(* IEC 61131-3 sources: daoli-st-library/DL_MathData (part 31) *)

(* ---- FC_DL_CalcDistance3D.st ---- *)
(*==============================================================================
 * 组件名称 (Component)  : FC_DL_CalcDistance3D
 * 所属子库 (Sublibrary) : DL_MathData
 * 当前版本 (Version)    : 1.0.0
 * 分类     (Category)   : 几何计算函数（Function · Math / Pure function）
 * 兼容性   (Platform)   : CODESYS 3.5 / TwinCAT 3 / 汇川 InoProShop / Machine Expert
 *                         仅依赖 Standard.library（SQRT / ABS / MAX），零厂商方言
 * 功能描述 (Function)   : 计算两点之间的三维欧氏距离，附带非有限值防护、
 *                         大数溢出缩放保护与三个分量差诊断输出。
 *                         平面（二维）距离不另设组件：把两个端点的 Z 坐标
 *                         同时填 0.0 即为其退化情形，规格明确禁止为凑数拆变体。
 *                         全程无内部状态，可任意频次调用。
 *
 * 【引脚契约 / Pin contract】
 *   输入 fX1 / fY1 / fZ1 : REAL — 点 1 的 X / Y / Z 坐标 [mm]，量程 ±1.0E6，
 *                                  平面场景把两个 Z 都填 0.0；
 *   输入 fX2 / fY2 / fZ2 : REAL — 点 2 的 X / Y / Z 坐标 [mm]，量程同上；
 *   输出 bValid          : BOOL — 六个输入全部有限（非 NaN、非无穷）= TRUE；
 *   输出 bSaturated      : BOOL — 本次计算进入大数缩放分支（结果仍然有效，
 *                                  但已落在置信区间，提示调用方复核量纲）；
 *   输出 fDeltaX/Y/Z     : REAL — 三个分量差 [mm]，便于现场诊断「差在哪个轴」；
 *   输出 uErrorId        : UDINT — 事件码，0 = 无。本件全部码为信息级。
 *   返回  值             : REAL — 距离 [mm]，恒非负；输入非法时返回 0.0。
 *
 * 【算法分步 / Algorithm steps（写死，防实现漂移）】
 *   ① 有限性闸门：六个输入任一非有限 → bValid FALSE、返回 0.0、置 0122 后早退。
 *      刻意**不返回 NaN**：NaN 会沿调用链污染下游滤波、比较与统计（历史教训）；
 *   ② 分量差：dX = X2 − X1（同 Y、Z），同时作为诊断输出；
 *   ③ 比例因子：fScale = MAX(|dX|, |dY|, |dZ|)，取最大分量作为量级基准；
 *   ④ 分支一（常规）：fScale 小于缩放阈值 → 直接 SQRT(dX² + dY² + dZ²)；
 *   ⑤ 分支二（缩放）：fScale 超阈值 → SQRT((dX/fScale)² + (dY/fScale)² +
 *      (dZ/fScale)²) × fScale。归一后每一项绝对值不超过 1，平方和不超过 3，
 *      彻底规避「大数先平方再开方」的中间溢出，结果为同一数学量的稳定写法；
 *   ⑥ 退化：三个分量差全为零（同一点）→ 返回 0.0 且不置任何码，因为距离为 0
 *      是合法结果而不是异常；
 *   ⑦ 后置守卫：最终结果非有限时（理论上不可达，防御性兜底）返回 0.0 并置 0122。
 *
 * 【数值安全 / Numeric safety】
 *   N1 非有限值用「区间比较取反」识别：NaN 参与任何有序比较均为假，故
 *      NOT(下限比较 AND 上限比较) 同时覆盖 NaN 与正负无穷，无需浮点判等；
 *   N2 缩放分支的分母恒大于阈值（阈值远大于 0），不存在除零；
 *   N3 平方和最多 3 项、每项不超过 1（缩放分支）或落在量程平方内（常规分支），
 *      不触碰 REAL 上界；
 *   N4 距离恒非负：SQRT 结果非负，早退路径返回 0.0，不存在负距离输出；
 *   N5 浮点判等红线：本件所有比较均为有序比较（小于 / 大于），唯一涉及「等于」
 *      的语义（同一点）由分量差与 0.0 做有序比较（小于容差）实现，不判等。
 *
 * 【边界防错清单 / Boundary guard list】
 *   B1 输入非有限（任一轴）→ bValid FALSE、返回 0.0、置 0122、不输出分量差；
 *   B2 两点重合 → 返回 0.0、bValid TRUE、bSaturated FALSE、零码（合法值）；
 *   B3 坐标取负 → 差值平方后符号消失，结果与全正坐标一致（V5 验证）；
 *   B4 量级超阈值 → 走缩放分支、bSaturated TRUE、置 0219（信息级，结果可用）；
 *   B5 结果非有限（兜底）→ 返回 0.0、置 0122，绝不把无穷扩散到调用方；
 *   B6 平面场景（Z 同值）→ 第三个分量差为 0，平方项为 0，公式自动退化，
 *      不需要任何分支判断，也不需要单独的二维入口。
 *
 * 【单位与量纲 / Units】
 *   输入输出统一按 [mm] 声明；若调用方用 [m] 或 [deg] 注入，输出随之为同单位，
 *   本件不做任何单位换算（换算属于标定层职责）。坐标差值超过 ±1.0E6 时
 *   结果仍然正确，但 bSaturated 会提示「已进入缩放置信区」，供质量追溯。
 *
 * 【与既有件的职责边界 / Family separation】
 *   FC_DL_PolygonArea       = 多点多边形面积与质心（面量）；
 *   FC_DL_LineIntersection  = 两条直线求交点（线量）；
 *   FB_DL_ElectronicCam /
 *   FB_DL_GantrySyncAxis    = 运动耦合，与几何距离无关；
 *   本件                    = 两点之间距离（点量），本族唯一的点对点度量件。
 *
 * 【调用示例 / Call example（仅行注释，不嵌套块注释）】
 *   // 视觉引导取料：料框中心与吸嘴当前坐标的三维距离，超过 50 mm 拒绝动作
 *   // fDist := FC_DL_CalcDistance3D(fX1 := fNozzleX, fY1 := fNozzleY, fZ1 := fNozzleZ,
 *   //          fX2 := fTargetX, fY2 := fTargetY, fZ2 := fTargetZ,
 *   //          bValid => bGeomOk, bSaturated => bGeomScaled,
 *   //          fDeltaX => fDx, fDeltaY => fDy, fDeltaZ => fDz,
 *   //          uErrorId => uGeomErr);
 *   // IF (NOT bGeomOk) OR (fDist > 50.0) THEN
 *   //     bMoveEnable := FALSE;
 *   // END_IF
 *
 * 【平台移植注意 / Porting notes】
 *   SQRT 为标准函数，输入非负时三平台行为一致；本件通过缩放分支保证 SQRT 的
 *   入参不会因中间溢出变成负值或无穷；阈值与容差全部来自 VAR CONSTANT，
 *   换平台不需要改动逻辑区任何一行。
 *
 * 【工程背景与应用场景 / Background and use cases】
 *   ① 视觉引导取料：吸嘴与目标点的三维偏差直接作为定位修正量；
 *   ② 三坐标 / 关节臂测点：两个测点之间的空间距离用于形位公差初筛；
 *   ③ 机器人安全距离：工具中心点与围栏采样点的距离，进入缩放区时提示复核；
 *   ④ 堆垛高度校核：料垛顶面采样点与理论平面的距离用于判定垛型合格。
 *
 * 【验收向量 / Acceptance vectors】
 *   V1 平面退化：(0, 0, 0) 到 (3, 4, 0) → 5.0（勾股 3-4-5）；
 *   V2 三维：(0, 0, 0) 到 (2, 3, 6) → 7.0（4 + 9 + 36 = 49，开方 7）；
 *   V3 同点：(1, 1, 1) 到 (1, 1, 1) → 0.0、bValid TRUE、零码；
 *   V4 非有限：fX1 为 NaN → 0.0、bValid FALSE、uErrorId 0122；
 *   V5 负坐标：(−3, −4, 0) 到 (0, 0, 0) → 5.0（差值绝对值参与平方）；
 *   V6 大数缩放：分量差 2.0E18 → bSaturated TRUE、uErrorId 0219、结果仍有限。
 *
 * 【事件码表 / Event code table（全部信息级，不置报警位）】
 *   16#0001_0122  输入含非有限值，返回 0.0 且 bValid 置假；
 *   16#0001_0219  模长超缩放阈值，已按缩放式求模，结果有效但进入置信区。
 *
 * 修订历史 (Revision)   :
 *   2026-11-15  v1.0.0  首版落盘（Round 11 · 泳道 A · LGF Math 组）
 *============================================================================*)
FUNCTION FC_DL_CalcDistance3D : REAL
VAR_INPUT
    fX1 : REAL;                            // 点 1 X 坐标 [mm]，量程 ±1.0E6 / Point 1 X coordinate [mm], range plus or minus 1.0E6
    fY1 : REAL;                            // 点 1 Y 坐标 [mm] / Point 1 Y coordinate [mm]
    fZ1 : REAL;                            // 点 1 Z 坐标 [mm]，平面场景填 0.0 / Point 1 Z coordinate [mm], 0.0 for planar use
    fX2 : REAL;                            // 点 2 X 坐标 [mm] / Point 2 X coordinate [mm]
    fY2 : REAL;                            // 点 2 Y 坐标 [mm] / Point 2 Y coordinate [mm]
    fZ2 : REAL;                            // 点 2 Z 坐标 [mm] / Point 2 Z coordinate [mm]
END_VAR
VAR_OUTPUT
    bValid     : BOOL;                     // 六个输入全为有限值 / All six inputs are finite
    bSaturated : BOOL;                     // 进入大数缩放分支 / The scaling branch was used
    fDeltaX    : REAL;                     // X 分量差 [mm]，诊断用 / X component delta [mm], for diagnostics
    fDeltaY    : REAL;                     // Y 分量差 [mm]，诊断用 / Y component delta [mm], for diagnostics
    fDeltaZ    : REAL;                     // Z 分量差 [mm]，诊断用 / Z component delta [mm], for diagnostics
    uErrorId   : UDINT;                    // 事件码，0 = 无 / Event code, 0 = none
END_VAR
VAR
    _fScale    : REAL;                     // 最大分量绝对值 [mm]，量级基准 / Largest absolute component [mm], magnitude basis
    _fSumSq    : REAL;                     // 归一后平方和 [-] / Normalised sum of squares
    _fResult   : REAL;                     // 距离工作副本 [mm] / Working copy of the distance [mm]
    _bFinite   : BOOL;                     // 有限性闸门标志 / Finiteness gate flag
END_VAR
VAR CONSTANT
    DL_FLOAT_EPS  : REAL  := 1.0E-6;       // 同点判定容差 [mm] / Coincident-point epsilon [mm]
    DL_INF_LIM    : REAL  := 1.0E37;       // 非有限值判据阈值，超此视为无穷 / Non-finite threshold, beyond is infinity
    DL_SCALE_THR  : REAL  := 1.0E18;       // 触发缩放的模长阈值 [mm] / Scaling threshold [mm]
    DL_DIST_ZERO  : REAL  := 0.0;          // 距离下界，恒非负 / Distance lower bound, never negative
    DL_ERR_NONFIN : UDINT := 16#0001_0122; // 输入非有限值的信息级码 / Info code for non-finite inputs
    DL_ERR_SCALED : UDINT := 16#0001_0219; // 已按缩放式求模的信息级码 / Info code for the scaled evaluation
END_VAR

(*------------------------------------------------------------------------------
 * 段 1｜返回值与输出预置（函数必须先给出安全返回值）
 *      Preset the return value and the outputs
 *   返回值预置 0.0：任何早退路径都带「无距离」语义，绝不返回 NaN 或未初始化值。
 *-----------------------------------------------------------------------------*)
FC_DL_CalcDistance3D := DL_DIST_ZERO;      // 返回值预置 0（Return preset to zero）
bValid     := TRUE;                        // 有效性预置通过（Validity preset to pass）
bSaturated := FALSE;                       // 缩放标志预置（Scaling flag preset）
fDeltaX    := DL_DIST_ZERO;                // 分量差预置 0（Delta X preset to zero）
fDeltaY    := DL_DIST_ZERO;                // 分量差预置 0（Delta Y preset to zero）
fDeltaZ    := DL_DIST_ZERO;                // 分量差预置 0（Delta Z preset to zero）
uErrorId   := 16#0000_0000;                // 事件码预清零（Event code preset to zero）
_bFinite   := TRUE;                        // 有限性闸门预置通过（Finiteness gate preset to pass）

(*------------------------------------------------------------------------------
 * 段 2｜有限性闸门（边界 B1 / 数值安全 N1）
 *      Finiteness gate over the six coordinates
 *   NaN 与任何有序比较的结果均为假，故「比较区间取反」同时覆盖 NaN 与无穷。
 *-----------------------------------------------------------------------------*)
IF NOT ((fX1 <= DL_INF_LIM) AND (fX1 >= -DL_INF_LIM)) THEN   // X1 非有限（X1 not finite）
    _bFinite := FALSE;                     // 闸门关闭（Close the gate）
END_IF
IF NOT ((fY1 <= DL_INF_LIM) AND (fY1 >= -DL_INF_LIM)) THEN   // Y1 非有限（Y1 not finite）
    _bFinite := FALSE;                     // 闸门关闭（Close the gate）
END_IF
IF NOT ((fZ1 <= DL_INF_LIM) AND (fZ1 >= -DL_INF_LIM)) THEN   // Z1 非有限（Z1 not finite）
    _bFinite := FALSE;                     // 闸门关闭（Close the gate）
END_IF
IF NOT ((fX2 <= DL_INF_LIM) AND (fX2 >= -DL_INF_LIM)) THEN   // X2 非有限（X2 not finite）
    _bFinite := FALSE;                     // 闸门关闭（Close the gate）
END_IF
IF NOT ((fY2 <= DL_INF_LIM) AND (fY2 >= -DL_INF_LIM)) THEN   // Y2 非有限（Y2 not finite）
    _bFinite := FALSE;                     // 闸门关闭（Close the gate）
END_IF
IF NOT ((fZ2 <= DL_INF_LIM) AND (fZ2 >= -DL_INF_LIM)) THEN   // Z2 非有限（Z2 not finite）
    _bFinite := FALSE;                     // 闸门关闭（Close the gate）
END_IF

IF NOT _bFinite THEN                       // 任一坐标不可判（Any coordinate undecidable）
    bValid   := FALSE;                     // 有效性置假（Validity cleared）
    uErrorId := DL_ERR_NONFIN;             // 置非有限值信息码（Raise the non-finite info code）
    RETURN;                                // 早退，返回值保持 0.0（Early exit, return stays zero）
END_IF

(*------------------------------------------------------------------------------
 * 段 3｜分量差计算（同时作为诊断输出，便于定位偏差轴）
 *      Component deltas, also exposed for diagnostics
 *-----------------------------------------------------------------------------*)
fDeltaX := fX2 - fX1;                      // X 分量差 [mm]（X delta）
fDeltaY := fY2 - fY1;                      // Y 分量差 [mm]（Y delta）
fDeltaZ := fZ2 - fZ1;                      // Z 分量差 [mm]（Z delta）

(*------------------------------------------------------------------------------
 * 段 4｜量级基准与分支选择（边界 B4 / 数值安全 N2）
 *      Magnitude basis and branch selection
 *   取最大分量绝对值作为量级基准：既用于同点判定，也用作缩放分母。
 *-----------------------------------------------------------------------------*)
_fScale := MAX(ABS(fDeltaX), MAX(ABS(fDeltaY), ABS(fDeltaZ)));  // 最大分量绝对值（Largest absolute component）

IF _fScale < DL_FLOAT_EPS THEN             // 三点差全在容差内，即同一点（Coincident points）
    FC_DL_CalcDistance3D := DL_DIST_ZERO;  // 同点距离为 0，属合法值（Zero distance, a legal result）
ELSIF _fScale <= DL_SCALE_THR THEN         // 常规量级，直接求模（Regular magnitude, direct evaluation）
    FC_DL_CalcDistance3D := SQRT(fDeltaX * fDeltaX
                               + fDeltaY * fDeltaY
                               + fDeltaZ * fDeltaZ);             // 直接平方和开方（Direct sum of squares）
ELSE                                       // 超阈值，走缩放分支（Above the threshold, scaled branch）
    _fResult := SQRT((fDeltaX / _fScale) * (fDeltaX / _fScale)
                   + (fDeltaY / _fScale) * (fDeltaY / _fScale)
                   + (fDeltaZ / _fScale) * (fDeltaZ / _fScale)) * _fScale;  // 归一平方和乘回量级（Normalised sum times the scale）
    FC_DL_CalcDistance3D := _fResult;      // 缩放结果（Scaled result）
    bSaturated := TRUE;                    // 置缩放标志（Raise the scaling flag）
    uErrorId   := DL_ERR_SCALED;           // 置缩放信息码（Raise the scaled info code）
END_IF

(*------------------------------------------------------------------------------
 * 段 5｜后置守卫（边界 B5 / 数值安全 N4）
 *      Post guard on the returned distance
 *   理论上不可达：缩放分支已把中间量限制在 3 以内，常规分支受量程约束。
 *   仍保留兜底，杜绝无穷或 NaN 扩散到调用方的滤波与比较链。
 *-----------------------------------------------------------------------------*)
IF NOT ((FC_DL_CalcDistance3D <= DL_INF_LIM) AND (FC_DL_CalcDistance3D >= -DL_INF_LIM)) THEN
    FC_DL_CalcDistance3D := DL_DIST_ZERO;  // 结果非有限，回退 0（Non-finite result, fall back to zero）
    bSaturated := FALSE;                   // 缩放标志复位（Scaling flag cleared）
    uErrorId   := DL_ERR_NONFIN;           // 置非有限值信息码（Raise the non-finite info code）
END_IF

IF FC_DL_CalcDistance3D < DL_DIST_ZERO THEN // 负距离不可能，兜底钳位（A negative distance is impossible）
    FC_DL_CalcDistance3D := DL_DIST_ZERO;  // 钳到 0，维持非负承诺（Clamp to zero, keep the non-negative promise）
END_IF
END_FUNCTION

(* ---- FC_DL_Crc8.st ---- *)
(*==============================================================================
 * 组件名称 (Component)  : FC_DL_Crc8
 * 所属子库 (Sublibrary) : DL_MathData
 * 归属目录 (Directory)  : C:\Library\DL_MathData
 * 当前版本 (Version)    : 1.0.0
 * 分类/来源标签         : 函数（FUNCTION）· 纯函数 · 参数化 8 位 CRC 校验
 *                         lgf-datahandling / oscat-network / crc8
 * 兼容性   (Platform)   : CODESYS 3.5 / TwinCAT 3 / 汇川 InoProShop / 施耐德
 *                         Machine Expert；仅用 Standard.library 的 SHL / XOR / AND
 *                         与显式枚举比较，不含查表常量数组，无实例依赖
 * 功能一句话 (Summary)  : 参数化 MSB-first 的 CRC-8 逐位算法，覆盖 ATM、SAE-J1850、
 *                         HITAG 三个变体，补齐本库 CRC 族的 8 位宽度。
 * 功能描述 (Function)   : 逐位算法，无查表、无状态、内存占用恒定。每个字节先与 CRC
 *                         寄存器异或，再做 8 次「看最高位、左移一位、条件异或多项式」，
 *                         全部字节处理完后与终值异或。三个变体只差多项式、初值、终值
 *                         三个参数，算法主体完全共用。典型现场用途：SMBus 与多数
 *                         传感器帧的 8 位校验、汽车与部分变频器状态帧的 SAE-J1850
 *                         校验、HITAG 类标签读写的同族变体、以及自定义短帧协议里
 *                         「厂家只给多项式、不给算法」时的快速对齐。
 * 与既有件边界 (Boundary): FC_DL_Crc16Modbus 做 16 位反射型、FC_DL_Crc32Ethernet 做
 *                         32 位、FC_DL_LrcChecksum 做纵向加和。本件只做 8 位且只做
 *                         MSB-first。反射型 8 位变体（多项式 16#31 的 MAXIM-DOW 一族）
 *                         位序相反，是另一套算法族，强行并入同一枚举会让「变体」概念
 *                         失真，故本件明确不立，留作后续独立件。
 * 三个变体参数表        :
 *   eCrc8Atm       多项式 16#07 初值 16#00 终值 16#00  典型 SMBus 与传感器帧
 *   eCrc8SaeJ1850  多项式 16#1D 初值 16#FF 终值 16#FF  典型汽车与变频器状态帧
 *   eCrc8Hitag     多项式 16#1D 初值 16#FF 终值 16#00  同族不同终值约定
 * 枚举映射表 (R31)      : eCrc8Atm 对应第 1 分支 ｜ eCrc8SaeJ1850 对应第 2 分支 ｜
 *                         eCrc8Hitag 对应第 3 分支 ｜ 其余脏值走兜底分支并回退 ATM。
 *                         三个合理值各有且仅有一个分支，兜底分支只接脏值。
 * 设计要点 (Key notes)  : ① 截断必须显式：入参长度超上限时先把截断标志置真，再把
 *                           实际参与长度改成上限，绝不静默按上限算却报「完整」；
 *                         ② 变体非法时回退到 ATM 而不是返回零：算一个可复算的值
 *                           便于现场与厂家的校验工具对表；
 *                         ③ 长度非法（小于 1）时直接返回零并置故障码，不进入循环；
 *                         ④ 纯函数：无内部状态、无跨周期残留，同入参同结果。
 *
 * 【验收向量 / Acceptance vectors（已按公开目录实算复核）】
 *   V1  ATM 标准串 9 字节（字符 1 到 9）→ 16#F4
 *   V2  SAE-J1850 同一串 → 16#4B
 *   V3  HITAG 同一串 → 16#B4
 *   V4  V-B 上限截断（R37 主向量）：nLen=200 → nProcessed=128、bTruncated=真、
 *       码 0141；不得静默按 128 算却报完整
 *   V5  V-A 域外：nLen=0 → 返回 16#00、码 0221、nProcessed=0、bTruncated=假
 *   V6  变体填 9（非法）→ 按 ATM 参数计算并置 0142，结果与 V1 相同
 *
 * 开源溯源 (Origin)     : 来源标签 lgf-datahandling 与 oscat-network。前者为免费闭源
 *                         发布的公开函数库手册，本件仅借鉴其数据处理组「校验按位宽
 *                         独立成族、CRC 家族参数化」的粒度事实；后者为 EPL-2.0 公开
 *                         库，本件仅借鉴「校验与诊断独立成族」的分类方式，未读取其
 *                         函数体。三个变体的多项式、初值、终值取自公开 CRC 参数目录
 *                         与各协议的公开规范，属公开常数。本件零代码行、零注释、
 *                         零数据结构引用，clean-room 独立实现，不构成衍生作品。
 * 码位说明 (Codes)      : 信息 16#0001_0141 长度已截断 ｜ 16#0001_0142 变体已回退
 *                         故障 16#0001_0221 长度非法。取号见本轮规格 §3.2。
 * 依赖说明 (Depends)    : 无 DL_ 内部依赖；仅 Standard.library 的 SHL / XOR / AND。
 * 镜像量清单 (R38)      : 本件无锁存副本，循环上界 nCount 由入口 nLen 一次导出后不再
 *                         读取入参，不存在锁存量与实时量混用面。
 * 红线自检 (Redline)    : 零全局变量表依赖 ｜ 零外部变量声明 ｜ 零物理地址直写
 *                         纯 IEC 61131-3 ｜ 无除法故无除零面 ｜ 循环上界全常量化
 *                         全变量与枚举项双语同行注释 ｜ 状态机 N/A（纯函数）
 * 修订历史 (Revision)   : 2026-11-15  v1.0.0  首版入库（Round 13 · 泳道 B CRC8 子族开族）
 *============================================================================*)

(*==============================================================================
 * 逐位算法推演 (Bitwise algorithm walk-through)：
 *   设寄存器初值 16#00、多项式 16#07，输入单字节 16#00
 *   第 1 步 寄存器异或字节后仍为 16#00
 *   第 2 步 连续 8 次「最高位为 0 则仅左移」，寄存器始终为 16#00
 *   终值与 16#00 异或后返回 16#00
 *   若输入为 16#80：异或后寄存器为 16#80，最高位为 1
 *   第 1 次移位得 16#00 再异或 16#07 得 16#07，其后 7 次移位按最高位判断继续推进
 *   可见「先判最高位、再移位、最后条件异或」的顺序不可颠倒，写反会得到另一族的
 *   校验值，且现象是「校验总是差一位固定值」，极难在总线上查出
 *============================================================================*)

(*==============================================================================
 * 调用示例 (Instance guide)：
 *   uCrc := FC_DL_Crc8(
 *              aData      := aFrame,
 *              nLen       := nLen,
 *              eVar       := E_DL_Crc8Variant.eCrc8Atm,
 *              nProcessed => nUsed,
 *              bTruncated => bCut,
 *              uErrorId   => uCode);
 *   提示：bCut 为真时说明帧长超出本件上限，校验值只覆盖前 128 字节，
 *         此时不得把它当作整帧校验结果使用。
 *============================================================================*)

TYPE E_DL_Crc8Variant :
(
    eCrc8Atm      := 0,  // SMBus 与多数传感器帧，多项式 16#07 初值 16#00 终值 16#00 / SMBus and most sensor frames
    eCrc8SaeJ1850 := 1,  // 汽车与部分变频器状态帧，多项式 16#1D 初值 16#FF 终值 16#FF / SAE J1850 flavour
    eCrc8Hitag    := 2   // 同族的另一终值约定，多项式 16#1D 初值 16#FF 终值 16#00 / HITAG flavour
);
END_TYPE

FUNCTION FC_DL_Crc8 : BYTE
VAR_INPUT
    aData : ARRAY[1..128] OF BYTE;                              // 数据缓冲区 [字节]，定长 128，未用位置填 0 / Data buffer, fixed 128 bytes, unused slots zeroed
    nLen  : INT;                                               // 有效字节数 [个]，域 1 到 128，超上限按截断规则处理 / Valid byte count, 1 to 128, truncated above the limit
    eVar  : E_DL_Crc8Variant := E_DL_Crc8Variant.eCrc8Atm;     // 变体选择 [枚举]，默认 ATM / Variant selector, ATM by default
END_VAR
VAR_OUTPUT
    nProcessed : INT;                                          // 实际参与计算的字节数 [个]，域 0 到 128 / Bytes actually processed, 0 to 128
    bTruncated : BOOL;                                         // 入参超上限被截断，截断发生时必须显式置真 / Set true explicitly whenever truncation happened
    uErrorId   : UDINT;                                        // 事件码，0 表示无事件 / Event code, zero means none
END_VAR
VAR
    uCrc    : BYTE;      // CRC 寄存器，逐位推进的运行值 [字节] / CRC register, the running value
    uPoly   : BYTE;      // 本次生效的多项式 [字节] / Effective polynomial
    uInit   : BYTE;      // 本次生效的初值 [字节] / Effective initial value
    uXorOut : BYTE;      // 本次生效的终值异或量 [字节] / Effective final xor value
    uByte   : BYTE;      // 当前处理字节快照 [字节] / Snapshot of the byte under processing
    nCount  : INT;       // 钳位后实际参与计算的字节数 [个] / Clamped byte count to process
    nI      : INT;       // 字节循环下标 [索引]，域 1 到 128 / Byte loop index, 1 to 128
    nBit    : INT;       // 位循环下标 [索引]，固定 1 到 8 / Bit loop index, fixed 1 to 8
    bMsb    : BOOL;      // 移位前最高位状态 [布尔] / Most significant bit state before the shift
    uCode   : UDINT;     // 码位暂存，出口单点写入 [码] / Code staging, written once at the exit
END_VAR
VAR CONSTANT
    DL_CRC8_MAXLEN : INT := 128;            // 定长上限 [字节]，与形参维度一致，避免大数组进栈 / Fixed upper bound matching the dimension
    DL_CRC8_BITS   : INT := 8;              // 每字节位循环次数 [次] / Bit iterations per byte
    DL_CRC8_MSB    : BYTE := 16#80;         // 最高位掩码 [位串] / Most significant bit mask
    DL_CRC8_MASK8  : BYTE := 16#FF;         // 八位满掩码，移位后裁掉溢出位 [位串] / Eight bit mask to drop the shifted out bit
    DL_CRC8_POLY_ATM : BYTE := 16#07;       // ATM 多项式 [字节] / ATM polynomial
    DL_CRC8_POLY_J1850 : BYTE := 16#1D;     // SAE-J1850 与 HITAG 多项式 [字节] / SAE J1850 and HITAG polynomial
    DL_CRC8_INIT_ATM : BYTE := 16#00;       // ATM 初值 [字节] / ATM initial value
    DL_CRC8_INIT_J1850 : BYTE := 16#FF;     // SAE-J1850 与 HITAG 初值 [字节] / SAE J1850 and HITAG initial value
    DL_CRC8_XOR_J1850 : BYTE := 16#FF;      // SAE-J1850 终值 [字节] / SAE J1850 final xor
    DL_CRC8_XOR_NONE : BYTE := 16#00;       // 无终值异或 [字节] / No final xor
END_VAR

(*------------------------------------------------------------------------------
 * 段 1｜安全预置：返回值落零，截断标志落假，码位落零
 *      Safe preset: zero return, truncation flag false, code cleared
 *      截断标志的初值必须是假，否则「恒真」与「从不置真」两种错误无法区分
 *      The flag starts false so that a stuck true and a never set true are distinguishable
 *-----------------------------------------------------------------------------*)
FC_DL_Crc8  := 16#00;
nProcessed  := 0;
bTruncated  := FALSE;
uErrorId    := 16#0000_0000;
uCode       := 16#0000_0000;
uCrc        := 16#00;
nCount      := 0;

(*------------------------------------------------------------------------------
 * 段 2｜长度闸门（边界 B1/B2）：小于 1 早退，大于上限先置截断标志再钳位
 *      Length gate: below one exits early, above the limit flags first then clamps
 *      顺序硬约束：先置标志、后改长度。反过来的写法会出现「已经按 128 算完、
 *      却因为标志被后面的赋值覆盖而报完整」的静默失真
 *      Order matters: flag first, then clamp, the reverse silently loses the evidence
 *-----------------------------------------------------------------------------*)
IF nLen < 1 THEN
    uErrorId := 16#0001_0221;   // 故障级：长度非法，返回零且不进入循环
    RETURN;
ELSIF nLen > DL_CRC8_MAXLEN THEN
    bTruncated := TRUE;         // 截断发生，先置标志
    nCount     := DL_CRC8_MAXLEN;
    uCode      := 16#0001_0141; // 信息级：已截断，实际只算前 128 字节
ELSE
    nCount := nLen;
END_IF

(*------------------------------------------------------------------------------
 * 段 3｜变体参数装载（边界 B3）：三个合法值逐一比较，脏值回退 ATM
 *      Variant parameter load: three legal values compared one by one, dirty falls back to ATM
 *      用等值列举而非区间判断：枚举底层是整数，区间判断会放过将来新增的成员
 *      Equality enumeration instead of a range test, a range would accept future members
 *-----------------------------------------------------------------------------*)
IF eVar = E_DL_Crc8Variant.eCrc8Atm THEN
    uPoly   := DL_CRC8_POLY_ATM;
    uInit   := DL_CRC8_INIT_ATM;
    uXorOut := DL_CRC8_XOR_NONE;
ELSIF eVar = E_DL_Crc8Variant.eCrc8SaeJ1850 THEN
    uPoly   := DL_CRC8_POLY_J1850;
    uInit   := DL_CRC8_INIT_J1850;
    uXorOut := DL_CRC8_XOR_J1850;
ELSIF eVar = E_DL_Crc8Variant.eCrc8Hitag THEN
    uPoly   := DL_CRC8_POLY_J1850;
    uInit   := DL_CRC8_INIT_J1850;
    uXorOut := DL_CRC8_XOR_NONE;
ELSE
    (* 兜底分支只接脏值：回退 ATM 参数并报信息级码，仍给出可复算的校验值 *)
    (* The fallback branch only sees dirty values, it falls back to ATM and reports *)
    uPoly   := DL_CRC8_POLY_ATM;
    uInit   := DL_CRC8_INIT_ATM;
    uXorOut := DL_CRC8_XOR_NONE;
    IF uCode = 16#0000_0000 THEN
        uCode := 16#0001_0142;
    END_IF
END_IF

(*------------------------------------------------------------------------------
 * 段 4｜逐字节、逐位计算（边界 B4/B5/B6）
 *      Byte-wise and bit-wise computation
 *      外层：nCount 已在段 2 保证 1 到 128，循环必执行且下标不越界
 *      内层：固定 8 次，顺序为「先取最高位、再左移、最后条件异或」
 *      移位后与满掩码相与，显式丢弃移出位，不依赖平台对 BYTE 移位的截断行为
 *-----------------------------------------------------------------------------*)
uCrc := uInit;

FOR nI := 1 TO nCount DO

    (* 写前下标双检，与形参维度 1 到 128 对齐 / Index double check against the declared dimension *)
    IF (nI >= 1) AND (nI <= DL_CRC8_MAXLEN) THEN

        uByte := aData[nI];
        uCrc  := uCrc XOR uByte;

        FOR nBit := 1 TO DL_CRC8_BITS DO
            bMsb := (uCrc AND DL_CRC8_MSB) <> 16#00;   // 步骤 1 移位前先捕获最高位
            uCrc := SHL(uCrc, 1) AND DL_CRC8_MASK8;    // 步骤 2 左移一位并裁掉溢出位
            IF bMsb THEN
                uCrc := uCrc XOR uPoly;               // 步骤 3 最高位为 1 时异或多项式
            END_IF
        END_FOR;

    END_IF

END_FOR;

(*------------------------------------------------------------------------------
 * 段 5｜终值异或与出口收口（边界 B7）
 *      Final xor and close out
 *-----------------------------------------------------------------------------*)
uCrc         := uCrc XOR uXorOut;
FC_DL_Crc8   := uCrc;
nProcessed   := nCount;
uErrorId     := uCode;      // 码位单点写入，全拍只写一次 / Single write point for the code
END_FUNCTION

(* ---- FC_DL_FactorialSat.st ---- *)
(*==============================================================================
 * 组件名称 (Component)  : FC_DL_FactorialSat
 * 所属子库 (Sublibrary) : DL_MathData
 * 当前版本 (Version)    : 1.0.1
 * 组件分类 (Category)   : 函数（FUNCTION）· 纯函数 · 阶乘（饱和输出）
 * 兼容性   (Platform)   : CODESYS 3.5 / TwinCAT 3 / 汇川 InoProShop / Schneider
 *                         Machine Expert；纯整数乘加，零浮点、零库依赖
 * 功能描述 (Function)   : 计算 n 的阶乘（n 为 0 到 12 的整数）。超出可算域时
 *                         饱和输出并置饱和标志与事件码，绝不返回错误数值冒充
 *                         结果。用于组合数与排列数、二项分布判定、配方阶乘
 *                         系数、多项式展开系数表初始化。
 * 可算域来源 (Why 12)   : 12 的阶乘等于 479001600，小于 DINT 上限 2147483647，
 *                         安全裕度约 4.5 倍；13 的阶乘等于 6227020800，已超
 *                         DINT 上限，故上限锁死在 12。若现场确需更大阶乘，
 *                         请改用 LINT 版本另立组件（不在本件内塞 MODE 参数）。
 * 设计要点 (Key notes)  : ① 饱和而非溢出：超域一律返回 12 的阶乘值并置 bSat，
 *                           调用方看 bSat 即知结果不可直接当真值使用；
 *                         ② 负入参约定：按 0 处理（0 的阶乘 = 1）并置 bSat 与
 *                           事件码，该约定在头注释与本段注释中双重写明，
 *                           避免现场把 1 误当正确答案；
 *                         ③ 累加器用 DINT，循环上界用钳位后的 nUsedN，
 *                           绝不用入参原值当循环上界；
 *                         ④ 无除法、无浮点、无不确定次数循环，故无需防死锁
 *                           计数器，也不需要浮点容差比较。
 * 开源溯源 (Origin)     : lgf-math。参考 LGF（Libre Graphical Framework）公开
 *                         函数库「Math」分类下阶乘函数的功能分类与参数域
 *                         （入参域 0 到 12、超域报错这一公开行为定义），只借
 *                         分类、参数域与该域约定，算法与实现 100% 自有
 *                         clean-room，不构成衍生作品。
 * 依赖     (Depends)    : 无 DL_ 内部依赖；无标准库功能块依赖
 * 故障码表 (Error codes):
 *   16#0001_011D【信息级】入参超域（负数或大于 12），饱和输出并置 bSat
 * 验收向量 (Acceptance) :
 *   V1 入参 0 → 1，bSat = FALSE
 *   V2 入参 5 → 120，bSat = FALSE
 *   V3 入参 12 → 479001600，bSat = FALSE
 *   V4 入参 13 → 479001600，bSat = TRUE，码 011D
 *   V5 入参 -3 → 1，bSat = TRUE，码 011D
 * 红线自检 (Redline)    : R1 零全局变量表与外部变量引用 ｜ R2 零物理地址直写
 *                         R3 纯 IEC 61131-3 ｜ R4 循环上界钳位、无除法故无除零面
 *                         R5 全变量中英双语同行注释 ｜ R6 N/A（纯函数无状态机）
 *                         R7 N/A（无实例调用）
 * 修订历史 (Revision)   :
 *   2026-11-15  v1.0.0  首版入库（Round 10 · Level 1 数学族回补）
 *   2026-11-15  v1.0.1  R10 终审修复（注释级）：R-FIX-1 累加器为 DINT 而循环
 *                       变量为 INT，原文 nAcc 乘 i 依赖隐式类型提升，违反
 *                       「不用隐式类型转换」红线（部分平台报隐式转换告警）；
 *                       改为显式 INT_TO_DINT。数值结果与全部验收向量不变。
 *============================================================================*)

(*==============================================================================
 * 阶乘查表基准 (Reference table，用于回归自检)：
 *   n    n!            与 DINT 上限之比
 *   0    1             可忽略
 *   1    1             可忽略
 *   2    2             可忽略
 *   3    6             可忽略
 *   4    24            可忽略
 *   5    120           可忽略
 *   6    720           可忽略
 *   7    5040          可忽略
 *   8    40320         可忽略
 *   9    362880        可忽略
 *   10   3628800       约千分之一点七
 *   11   39916800      约百分之一点九
 *   12   479001600     约百分之二十二
 *   13   6227020800    已超上限，本件拒绝并饱和到 12 的阶乘
 *   上表只用整数字面量，不含浮点，可逐条作为仿真回归的期望值。
 *============================================================================*)

(*==============================================================================
 * 算法推演 (Worked traces)：
 *   推演 1  入参 0
 *     段 2 非负，通过；段 3 不超上限，通过
 *     段 4 有效 n 取 0，累加器取 1
 *     循环从 2 到 0，起止倒置，一次都不执行，累加器仍为 1
 *     段 5 返回 1，饱和标志假
 *   推演 2  入参 5
 *     段 4 有效 n 取 5，累加器取 1
 *     循环依次乘 2、3、4、5，得 120
 *   推演 3  入参 12
 *     循环依次乘 2 到 12，终值 479001600，未溢出，饱和标志假
 *   推演 4  入参 13
 *     段 3 超上限成立，有效 n 钳到 12，饱和标志真，置码 011D
 *     立即返回饱和值，不进入循环（避免真的算出溢出数）
 *   推演 5  入参 负 3
 *     段 2 判负成立，按 0 处理并置饱和标志与码，返回 1
 *============================================================================*)

(*==============================================================================
 * 饱和语义与调用契约 (Contract)：
 *   1 饱和标志为假时，返回值可以当作数学上的精确阶乘直接参与后续整数运算；
 *   2 饱和标志为真时，返回值只是「可算域内最大的阶乘」，不具备数值意义，
 *     调用方必须把它当作「超出能力」的信号，不得继续参与运算；
 *   3 负入参按 0 处理是本库的显式约定：负数的阶乘在实数域无定义，
 *     返回 1 并置饱和标志，既避免了未定义行为，也让 HMI 有可显示的确定值；
 *   4 本件不抛异常、不阻塞、不依赖任何库，可在中断级任务中安全调用。
 *============================================================================*)

(*==============================================================================
 * 调用示例 (Instance guide)：
 *   组合数 C(n, k) 的分子计算（n 不超过 12，故可在本件域内完成）：
 *     nFac := FC_DL_FactorialSat(nValue := n);
 *     kFac := FC_DL_FactorialSat(nValue := k);
 *     nkFac := FC_DL_FactorialSat(nValue := n - k);
 *     IF (NOT bSat) AND (kFac > 0) AND (nkFac > 0) THEN
 *         nComb := nFac / (kFac * nkFac);
 *     END_IF
 *   注意：三个调用各自有独立的饱和标志，必须全部为假才可继续；只判其中
 *   一个是现场最常见的越域漏检，会在组合数上产生数量级错误。
 *============================================================================*)

(*==============================================================================
 * 与相关件的关系 (Related components)：
 *   1 本件只负责阶乘，不做组合数与排列数；组合数需要三次阶乘再相除，由
 *     调用方按上节示例组合，本库不提供「组合数巨无霸块」；
 *   2 阶乘与幂运算是两回事：本件不做幂，任意次幂请按幂律自行乘算或改用
 *     对数法，切勿用阶乘近似幂；
 *   3 本件的饱和语义与 FB_DL_PresetCounterSat 的饱和语义同源（都是「到边界
 *     即停并给标志」），但二者管辖对象不同，不得互相替代。
 *============================================================================*)

(*==============================================================================
 * 类型与容量说明 (Type capacity)：
 *   入参 nValue 用 INT，是因为可算域只有 0 到 12，用 DINT 会误导调用方以为
 *   能算更大；返回值用 DINT，是因为 12 的阶乘已经接近三十二位有符号上限的
 *   四分之一，再用 INT 会溢出。二者刻意不同，请勿「统一类型」后重写。
 *   若现场确需 13 以上的阶乘，请另立 LINT 版本组件，本件不扩域。
 *============================================================================*)

(*==============================================================================
 * 执行代价与扫描时间 (Cost)：
 *   最坏路径是入参 12，循环体执行十一次整数乘法，在任何一款目标 PLC 上都
 *   只占纳秒到微秒量级，可以放心放在每毫秒中断任务里调用；但若在单次扫描
 *   里对同一组数据反复调用上百次（例如批量初始化系数表），请先把结果缓存
 *   到数组里，不要每拍重算——省下的不是乘法时间，而是调用开销与代码体积。
 *   本件不含除法、不含浮点、不含不定次数循环，故最坏执行时间可静态界定，
 *   满足硬实时任务对最长执行路径可证明的要求。
 *============================================================================*)

FUNCTION FC_DL_FactorialSat : DINT
VAR_INPUT
    nValue : INT := 0;       // 自然数 n，有效域 0 到 12，负数按 0 处理 [无量纲] / Natural number, valid 0 to 12, negatives treated as zero
END_VAR
VAR_OUTPUT
    bSat     : BOOL;         // 饱和标志：入参超域或结果溢出为 TRUE [-] / TRUE when the input is out of domain or saturated
    nUsedN   : INT;          // 实际参与计算并钳位后的 n [无量纲] / Effective n after clamping
    uErrorId : UDINT;        // 事件码，0 = 无事件 / Event code, 0 = no event
END_VAR
VAR
    i    : INT;              // 循环索引，域 2 到 nUsedN [无量纲] / Loop index, 2 to nUsedN
    nAcc : DINT;             // 累加器，12 的阶乘不溢出 [无量纲] / Accumulator, twelve factorial never overflows
END_VAR
VAR CONSTANT
    DL_FACT_MAX_N : INT  := 12;         // 最大可算 n，13 的阶乘已超 DINT 上限 [无量纲] / Highest computable n
    DL_FACT_SAT   : DINT := 479001600;  // 饱和输出值，等于 12 的阶乘 [无量纲] / Saturation output, twelve factorial
    DL_FACT_ZERO  : DINT := 1;          // 0 的阶乘定义值 [无量纲] / Zero factorial by definition
    DL_FACT_BASE  : INT  := 2;          // 循环起点，1 的阶乘无需乘算 [无量纲] / Loop start index
END_VAR

(*------------------------------------------------------------------------------
 * 段 1｜输出与返回值预置
 *      Pre-set outputs and return value
 *-----------------------------------------------------------------------------*)
FC_DL_FactorialSat := DL_FACT_ZERO;
bSat     := FALSE;
nUsedN   := 0;
uErrorId := 16#0000_0000;

(*------------------------------------------------------------------------------
 * 段 2｜负入参（边界 B1）：按 0 处理并置饱和
 *      Negative input (boundary B1): treated as zero and flagged saturated
 *      约定写明：负数返回 1（等于 0 的阶乘）且 bSat 为 TRUE，调用方必须看标志
 *-----------------------------------------------------------------------------*)
IF nValue < 0 THEN
    nUsedN            := 0;
    bSat              := TRUE;
    uErrorId          := 16#0001_011D;
    FC_DL_FactorialSat := DL_FACT_ZERO;
    RETURN;
END_IF

(*------------------------------------------------------------------------------
 * 段 3｜超上限入参（边界 B2）：饱和到 12 的阶乘
 *      Input above the upper bound (boundary B2): saturate to twelve factorial
 *-----------------------------------------------------------------------------*)
IF nValue > DL_FACT_MAX_N THEN
    nUsedN            := DL_FACT_MAX_N;
    bSat              := TRUE;
    uErrorId          := 16#0001_011D;
    FC_DL_FactorialSat := DL_FACT_SAT;
    RETURN;
END_IF

(*------------------------------------------------------------------------------
 * 段 4｜主路径：从 2 连乘到 n，循环上界只用钳位后的 nUsedN
 *      Main path: multiply from two up to n, the bound is the clamped value
 *-----------------------------------------------------------------------------*)
nUsedN := nValue;
nAcc   := DL_FACT_ZERO;

FOR i := DL_FACT_BASE TO nUsedN DO
    nAcc := nAcc * INT_TO_DINT(i);   // 显式升位：INT 乘 DINT 的隐式转换在部分平台告警
END_FOR

(*------------------------------------------------------------------------------
 * 段 5｜合法收口：bSat 为 FALSE 时调用方可直接当精确值使用（契约级承诺）
 *      Legal close-out: with bSat FALSE the value is exact by contract
 *-----------------------------------------------------------------------------*)
FC_DL_FactorialSat := nAcc;
END_FUNCTION

(* ---- FC_DL_Matrix3Inverse.st ---- *)
(*==============================================================================
 * 组件名称 (Component)  : FC_DL_Matrix3Inverse
 * 所属子库 (Sublibrary) : DL_MathData
 * 归属目录 (Directory)  : C:\Library\DL_MathData
 * 当前版本 (Version)    : 1.0.1
 * 分类/来源标签         : 函数（FUNCTION）· 纯函数 · 三阶方阵求逆
 *                         lgf-math / matrix / affine-transform
 * 兼容性   (Platform)   : CODESYS 3.5 / TwinCAT 3 / 汇川 InoProShop / 施耐德
 *                         Machine Expert；仅用 Standard.library 的 ABS / MIN /
 *                         MAX / LIMIT，无矩阵库依赖，无循环嵌套
 * 功能一句话 (Summary)  : 3 乘 3 实数矩阵按伴随矩阵法解析求逆，含相对奇异判据与
 *                         出口夹域，失败时逆矩阵整体置 0 且绝不输出非数。
 * 功能描述 (Function)   : 九个元素行主序传入，先用余子式展开算行列式，再用伴随矩阵
 *                         除以行列式得到逆。全过程为定长表达式，无主元选取、无嵌套
 *                         循环、无分支跳步，因此同一输入在同一平台上的每一步中间量
 *                         都可复算。典型现场用途：视觉与机器人手眼标定的反解、仿射
 *                         变换的逆映射（像素坐标反算机械坐标）、三传感器三角定位的
 *                         线性方程组求解、标定矩阵在校验工位上的逐拍复核。
 * 为什么不用高斯消元    : 三阶的解析逆是固定九个表达式，无分支、无主元交换、无循环，
 *                         天然满足「纯函数、确定性、可逐拍复算」三条验收要求；高斯
 *                         消元需要三层嵌套循环加主元选择分支，在三阶规模上没有任何
 *                         数值或性能收益，却引入了「主元为 0 时要换行」的分支面。
 * 数值判据（本件关键）  : 不用绝对阈值判奇异。矩阵元素量纲相差一千倍时（毫米级标定
 *                         矩阵与微米级标定矩阵），绝对阈值必然失效：同一个 1.0E-9 的
 *                         绝对门槛对前者过严、对后者过松。本件改用相对判据
 *                         「行列式绝对值 小于等于 相对容差 乘 最大元素绝对值的立方」，
 *                         于是同一个相对容差在两种量纲下都成立。fDetEps 是相对量，
 *                         默认 1.0E-9，不是绝对量，切勿按绝对行列式理解。
 * 与既有件边界 (Boundary): FC_DL_LineIntersection 解两直线交点、FC_DL_CalcDistance3D 算
 *                         点距、FC_DL_PolygonArea 算多边形面积。三者都是定式几何量；
 *                         本件提供通用可逆性判定与逆矩阵，供标定与坐标变换链复用。
 *                         矩阵子族从此件开族，后续四阶与伪逆另立。
 * 设计要点 (Key notes)  : ① 入口先做非有限元素体检：任一元为无穷或非数则整件拒绝，
 *                           而不是让脏值流进行列式把九个输出全污染；
 *                         ② 相对奇异判据只用「行列式、最大元素绝对值、相对容差」
 *                           三个量，判据、守卫、封顶三者同向（见下方三元一致表）；
 *                         ③ 除法前显式确认行列式非零，即使奇异判据已保证；
 *                         ④ 出口夹域：每个逆元素先判有限再夹进上下界，失败路径整体
 *                           置 0 而不置非数，上层拿到的是「明确不可信」而不是毒值；
 *                         ⑤ 纯函数：无内部状态、无跨周期残留，同入参同结果。
 *
 * 【三元一致表 / Guard and criterion consistency (R35)】
 *   守卫：最大元素绝对值 fMaxAbs 仅用于构造立方尺度，不做封顶
 *   封顶：奇异性阈值等于 相对容差 乘 fMaxAbs 的立方，阈值随量纲自动缩放
 *   判据：行列式绝对值 小于等于 该阈值 即判奇异，与守卫同向，无「守卫通过但判据更宽」的缝
 *
 * 【验收向量 / Acceptance vectors】
 *   V1  单位阵 → 逆等于自身、行列式 1.0、返回真
 *   V2  对角阵「2 4 5」→ 逆为对角「0.5 0.25 0.2」、行列式 40.0、返回真
 *   V3  V-A 奇异专测：第一行「1 2 3」、第二行「2 4 6」（第二行是第一行两倍）、
 *       第三行「7 8 9」→ 行列式 0、返回假、码 0225、逆矩阵全 0
 *   V4  V-B 相对判据专测：V3 整体乘 1.0E-6 → 行列式量级 1.0E-18，绝对阈值必然
 *       误判为可逆；本件按相对判据仍返回假、码 0225（此向量是本判据存在的唯一理由）
 *   V5  V-D 出口夹域：任一元素传入非数 → 码 014B、返回假、逆矩阵全 0（不输出非数）
 *   V6  V-D 相对容差非法：相对容差传 0 → 码 014C、按默认 1.0E-9 继续，返回真
 *   V7  病态提示：对角阵「1 1 1.0E-6」且相对容差取 1.0E-12 → 条件数粗估
 *       fCondEst = |det| 除 maxAbs 立方 = 1.0E-6 除 1 = 1.0E-6（v1.0.1 勘误，
 *       旧版误记 1.0E-18），落在「超 10 倍容差、低于 1.0E-3」区间内，
 *       逆已给出、码 014A（提示精度不保）
 *
 * 开源溯源 (Origin)     : 来源标签 lgf-math。LGF（Libre Graphical Framework）为免费
 *                         闭源发布的公开函数库手册，本件仅借鉴其数学组存在「矩阵」
 *                         子族（含求逆、转置、乘加等按阶数分件的粒度事实），作为
 *                         子族开族的立项依据；许可证按其发布方条款仅作分类参考。
 *                         伴随矩阵法与余子式展开属公开线性代数经典内容，本件零代码行、
 *                         零注释、零数据结构引用，clean-room 独立实现，不构成衍生作品。
 * 码位说明 (Codes)      : 信息 16#0001_014A 病态但已给逆 ｜ 16#0001_014B 含非有限元素
 *                         16#0001_014C 相对容差非正已用默认
 *                         故障 16#0001_0225 矩阵奇异。取号见本轮规格 §3.2，
 *                         与定长串子族 0143 到 0149 不重叠。
 * 依赖说明 (Depends)    : 无 DL_ 内部依赖；仅 Standard.library 的 ABS / LIMIT。
 * 镜像量清单 (R38)      : 无锁存副本。九个元素入口一次拷入局部数组，其后全部表达式
 *                         只用局部数组与入口标量，不再读形参数组，故调用方在本件返回前
 *                         改写入参数组也不会撕裂中间量。
 * 偏离留档 (Deviation)  : 形参数组维度用字面量 9（行主序九个元素），逻辑区用常量
 *                         DL_M3_CNT 表达同一上界，二者字面一致，不构成双源。
 * 红线自检 (Redline)    : 零全局变量表依赖 ｜ 零外部变量声明 ｜ 零物理地址直写
 *                         纯 IEC 61131-3 ｜ 每处除法前判行列式非零 ｜ 浮点不用等值比较
 *                         全变量双语同行注释 ｜ 状态机 N/A（纯函数）｜ 无定时器实例
 * 修订历史 (Revision)   : 2026-11-15  v1.0.0  首版入库（Round 13 · 泳道 B 矩阵子族开族）
 *                         2026-11-16  v1.0.1  终审勘误：验收向量 V7 的条件数粗估值由
 *                         误记的 1.0E-18 更正为实算值 1.0E-6（fCondEst = |det| 除
 *                         maxAbs 立方），仅更正头注释记载，判定逻辑与码位不变
 *============================================================================*)

(*==============================================================================
 * 行主序排布与余子式对应 (Row-major layout)：
 *   元素 1 到 3 是第一行，4 到 6 是第二行，7 到 9 是第三行
 *   行列式按第一行展开，三个余子式分别用第二三两行的元素组合
 *   伴随矩阵是余子式矩阵的转置，故逆矩阵第 2 个元素用的是「第 1 行第 2 列」的
 *   代数余子式，而不是第 2 行第 1 列的，写反会让逆矩阵整体转置
 *   对角阵是最容易验证排布是否写反的例子：转置后仍然是对角阵，看不出错，
 *   所以验收向量必须包含非对角元素非零的矩阵（V3 的三行两两不成比例）
 *============================================================================*)

FUNCTION FC_DL_Matrix3Inverse : BOOL
VAR_INPUT
    afM     : ARRAY[1..9] OF LREAL;   // 行主序 3 乘 3 矩阵 [无量纲或工程单位] / Row-major three by three matrix
    fDetEps : LREAL := 1.0E-9;        // 相对奇异判据 [无量纲]，非正时按默认处理 / Relative singularity epsilon, defaulted when not positive
END_VAR
VAR_OUTPUT
    afInv   : ARRAY[1..9] OF LREAL;   // 逆矩阵，行主序，失败时全 0 [无量纲或工程单位] / Inverse in row-major order, zeroed on failure
    fDet    : LREAL;                  // 行列式值 [无量纲或工程单位立方] / Determinant value
    fCondEst: LREAL;                  // 条件数粗估，越小越病态 [无量纲] / Coarse condition estimate, smaller means worse
    uErrorId: UDINT;                  // 事件码，0 表示无事件 / Event code, zero means none
END_VAR
VAR
    aV      : ARRAY[1..9] OF LREAL;   // 入参局部副本，非有限元素已按 0 落盘 [无量纲] / Local copy with non-finite elements zeroed
    aW      : ARRAY[1..9] OF LREAL;   // 伴随矩阵九个分子，尚未除以行列式 [无量纲] / Nine adjugate numerators before the division
    fMaxAbs : LREAL;                  // 九个元素绝对值的最大值 [同元素单位] / Largest absolute element
    fScale  : LREAL;                  // 最大元素绝对值的立方，作相对尺度的分母 [同元素单位立方] / Cube of the largest absolute element
    fDetR   : LREAL;                  // 行列式计算值 [同元素单位立方] / Computed determinant
    fCofA   : LREAL;                  // 第一行第一列余子式 [同元素单位平方] / First cofactor
    fCofB   : LREAL;                  // 第一行第二列余子式 [同元素单位平方] / Second cofactor
    fCofC   : LREAL;                  // 第一行第三列余子式 [同元素单位平方] / Third cofactor
    fEps    : LREAL;                  // 本次生效的相对容差 [无量纲] / Effective relative epsilon
    fThresh : LREAL;                  // 奇异性阈值，等于容差乘尺度 [同元素单位立方] / Singularity threshold
    fTmp    : LREAL;                  // 逆元素中间量 [无量纲] / Inverse element intermediate
    nI      : INT;                    // 元素循环下标 [索引]，1 到 9 / Element loop index, 1 to 9
    bNonFin : BOOL;                   // 含非有限元素标记 / Non-finite element flag
    uCode   : UDINT;                  // 码位暂存，出口单点写入 [码] / Code staging, written once at the exit
END_VAR
VAR CONSTANT
    DL_M3_CNT      : INT := 9;              // 元素个数 [个]，与形参维度一致 / Element count, matches the dimension
    DL_M3_FINITE   : LREAL := 1.0E308;      // 有限性上界 [无量纲]，用于拦无穷与非数 / Finiteness bound
    DL_M3_CONDWARN : LREAL := 1.0E-3;       // 病态提示门限 [无量纲]，小于此值提示精度不保 / Ill-conditioned warning threshold
    DL_M3_CONDK    : LREAL := 10.0;         // 病态提示的相对倍数 [无量纲] / Multiplier for the ill-conditioned test
    DL_M3_EPSDEF   : LREAL := 1.0E-9;       // 默认相对容差 [无量纲] / Default relative epsilon
END_VAR

(*------------------------------------------------------------------------------
 * 段 1｜输出预置（边界 B1，R43）：失败路径的逆矩阵必须是全 0，不是全非数
 *      Pre-set: the failure path publishes all zeros, never not-a-number values
 *      逐元素预置而不是整块赋值，保证每一路出口都在声明域内
 *      Element by element, so every exit path stays inside the declared domain
 *-----------------------------------------------------------------------------*)
FC_DL_Matrix3Inverse := FALSE;
FOR nI := 1 TO DL_M3_CNT DO
    afInv[nI] := 0.0;
    aV[nI]    := 0.0;
    aW[nI]    := 0.0;
END_FOR;
fDet      := 0.0;
fCondEst  := 0.0;
uErrorId  := 16#0000_0000;
uCode     := 16#0000_0000;
fMaxAbs   := 0.0;
fScale    := 0.0;
fDetR     := 0.0;
fThresh   := 0.0;
bNonFin   := FALSE;

(*------------------------------------------------------------------------------
 * 段 2｜相对容差闸门（边界 B2）：非正容差退回默认，不阻断计算
 *      Epsilon gate: a non-positive epsilon falls back to the default
 *      容差为 0 会让所有矩阵都判奇异，为负更无意义；退回默认并报信息级码
 *      A zero epsilon would mark every matrix singular, so the default is used
 *-----------------------------------------------------------------------------*)
IF fDetEps > 0.0 THEN
    fEps := fDetEps;
ELSE
    fEps    := DL_M3_EPSDEF;
    uCode   := 16#0001_014C;
END_IF

(*------------------------------------------------------------------------------
 * 段 3｜非有限元素体检（边界 B3）：任一元为无穷或非数则整件拒绝
 *      Non-finite check: a single bad element rejects the whole call
 *      体检式：两个比较同时成立才算有限，非数会让两个比较都为假，故此式一并拦截
 *      Both comparisons must hold, a not-a-number fails both and is caught
 *      脏值按 0 落进副本仅用于让码位与诊断可读，本路径不会继续求逆
 *      The dirty value is stored as zero only so the diagnostics stay readable
 *-----------------------------------------------------------------------------*)
FOR nI := 1 TO DL_M3_CNT DO
    IF (afM[nI] <= DL_M3_FINITE) AND (afM[nI] >= -DL_M3_FINITE) THEN
        aV[nI] := afM[nI];
    ELSE
        aV[nI]    := 0.0;
        bNonFin   := TRUE;
    END_IF
END_FOR;

IF bNonFin THEN
    uErrorId := 16#0001_014B;   // 信息级：含非有限元素，逆矩阵保持全 0
    RETURN;
END_IF

(*------------------------------------------------------------------------------
 * 段 4｜相对尺度（边界 B4）：九个元素绝对值的最大值，其立方即量纲尺度
 *      Relative scale: the largest absolute element, its cube is the scale
 *      尺度为零意味着整张矩阵全零，后续阈值也为零，行列式零必然被判奇异
 *      A zero scale means an all zero matrix, the threshold collapses to zero as well
 *-----------------------------------------------------------------------------*)
FOR nI := 1 TO DL_M3_CNT DO
    IF ABS(aV[nI]) > fMaxAbs THEN
        fMaxAbs := ABS(aV[nI]);
    END_IF
END_FOR;

fScale := fMaxAbs * fMaxAbs * fMaxAbs;

(*------------------------------------------------------------------------------
 * 段 5｜行列式与条件数粗估（边界 B5）：按第一行展开，三个余子式先行
 *      Determinant and condition estimate: expand along the first row
 *      除法前的显式判零放在段 7，此处只算不除
 *      No division here, the guarded division lives in stage seven
 *-----------------------------------------------------------------------------*)
fCofA := aV[5] * aV[9] - aV[6] * aV[8];   // 第一行第一列余子式 / Cofactor of row one column one
fCofB := aV[4] * aV[9] - aV[6] * aV[7];   // 第一行第二列余子式 / Cofactor of row one column two
fCofC := aV[4] * aV[8] - aV[5] * aV[7];   // 第一行第三列余子式 / Cofactor of row one column three

fDetR := aV[1] * fCofA - aV[2] * fCofB + aV[3] * fCofC;

IF (fDetR <= DL_M3_FINITE) AND (fDetR >= -DL_M3_FINITE) THEN
    fDet := fDetR;                          // 有限才发布，否则保持 0 / Published only when finite
ELSE
    fDet := 0.0;
END_IF

fCondEst := 0.0;
IF fScale > 0.0 THEN
    fTmp := ABS(fDetR) / fScale;            // 除数是正数，无除零面
    IF (fTmp <= DL_M3_FINITE) AND (fTmp >= -DL_M3_FINITE) THEN
        fCondEst := fTmp;
    ELSE
        fCondEst := 0.0;
    END_IF
END_IF

(*------------------------------------------------------------------------------
 * 段 6｜相对奇异判定（边界 B6）：阈值随量纲缩放，判据与守卫同向
 *      Relative singularity test: the threshold scales with the magnitude
 *      阈值等于容差乘尺度；全零矩阵时尺度与阈值同为 0，判据「0 小于等于 0」成立
 *      With an all zero matrix both sides collapse to zero and the test still holds
 *-----------------------------------------------------------------------------*)
fThresh := fEps * fScale;

IF ABS(fDetR) <= fThresh THEN
    uErrorId := 16#0001_0225;   // 故障级：奇异，逆不可得，逆矩阵保持全 0
    RETURN;
END_IF

(*------------------------------------------------------------------------------
 * 段 7｜伴随矩阵与除法（边界 B7）：先显式确认行列式非零，再逐元素相除
 *      Adjugate and division: confirm a non-zero determinant before dividing
 *      奇异判据已保证行列式非零，此处仍显式判一次，属于除零面的第二道锁
 *      The singularity test already guarantees it, this is the second lock
 *-----------------------------------------------------------------------------*)
IF (fDetR > 0.0) OR (fDetR < 0.0) THEN

    aW[1] := aV[5] * aV[9] - aV[6] * aV[8];
    aW[2] := aV[3] * aV[8] - aV[2] * aV[9];
    aW[3] := aV[2] * aV[6] - aV[3] * aV[5];
    aW[4] := aV[6] * aV[7] - aV[4] * aV[9];
    aW[5] := aV[1] * aV[9] - aV[3] * aV[7];
    aW[6] := aV[3] * aV[4] - aV[1] * aV[6];
    aW[7] := aV[4] * aV[8] - aV[5] * aV[7];
    aW[8] := aV[2] * aV[7] - aV[1] * aV[8];
    aW[9] := aV[1] * aV[5] - aV[2] * aV[4];

    FOR nI := 1 TO DL_M3_CNT DO
        fTmp := aW[nI] / fDetR;
        (* 出口夹域：非有限先归零，再夹进上下界，出口值必在声明域内 *)
        (* Exit clamp: non-finite collapses to zero, then everything is bounded *)
        IF (fTmp <= DL_M3_FINITE) AND (fTmp >= -DL_M3_FINITE) THEN
            afInv[nI] := LIMIT(-DL_M3_FINITE, fTmp, DL_M3_FINITE);
        ELSE
            afInv[nI] := 0.0;
        END_IF
    END_FOR;

ELSE

    uErrorId := 16#0001_0225;   // 兜底：行列式恰为零，与奇异判据同码
    RETURN;

END_IF

(*------------------------------------------------------------------------------
 * 段 8｜病态提示与成功收口（边界 B8）
 *      Ill-conditioning notice and the success close out
 *      条件数粗估小于千分之一但明显高于容差，说明逆虽给出、精度不保
 *      Below one thousandth yet well above the epsilon, the inverse is shown but shaky
 *-----------------------------------------------------------------------------*)
IF (fCondEst < DL_M3_CONDWARN) AND (fCondEst > (DL_M3_CONDK * fEps)) THEN
    uCode := 16#0001_014A;      // 信息级：病态，逆已给出
END_IF

uErrorId := uCode;              // 码位单点写入，全拍只写一次
FC_DL_Matrix3Inverse := TRUE;
END_FUNCTION

(* ---- FC_DL_NthRoot.st ---- *)
(*==============================================================================
 * 组件名称 (Component)  : FC_DL_NthRoot
 * 所属子库 (Sublibrary) : DL_MathData
 * 当前版本 (Version)    : 1.0.0
 * 组件分类 (Category)   : 函数（FUNCTION）· 纯函数 · N 次方根（奇偶次分治）
 * 兼容性   (Platform)   : CODESYS 3.5 / TwinCAT 3 / 汇川 InoProShop / Schneider
 *                         Machine Expert；仅用 Standard.library 的 EXP / LN /
 *                         SQRT / ABS，无任何厂商私有数学库锁定
 * 功能描述 (Function)   : 计算 x 的 n 次方根（x 的 1 除以 n 次幂）。标准库只有
 *                         SQRT（二次方根），本件补齐任意次根，覆盖几何平均、
 *                         等效值折算、按幂律反算（泵与风机相似定律反算转速比、
 *                         面积等效直径、均方根到峰值折算）等场景。
 * 与既有件边界 (Boundary): 本库无同类件；FC_DL_LinearScale 与
 *                         FC_DL_MultiPointLinear 是线性与折线映射，与幂运算
 *                         无语义交集，不得互相替代。
 * 设计要点 (Key notes)  : ① 奇偶分治是负数的唯一正确解：偶次根在实数域无解，
 *                           必须拒绝并给码，绝不能返回绝对值的结果冒充；
 *                           奇次根取绝对值求根后取反，符号必须保留；
 *                         ② 零与近零直接返回 0，绕开 LN(0) 的负无穷陷阱；
 *                         ③ 二次根特判走 SQRT，精度优于对数法；一次根特判
 *                           直接返回原值；底数为 1 特判省一次 EXP / LN；
 *                         ④ 对数法用 EXP(LN(绝对值) 除以 n)，除数恒大于等于 1
 *                           （已由根次数域校验保证），无除零面；
 *                         ⑤ 结果有限性复检：EXP 在极端入参下可能溢出为非有限值，
 *                           必须复检后置 bValid，绝不把无穷大当结果交出去；
 *                         ⑥ 明确禁用迭代牛顿法：收敛次数不定，违反 PLC 的确定性
 *                           时间约束，现场表现为「同一入参偶尔多占一个周期」。
 * 开源溯源 (Origin)     : lgf-math。参考 LGF（Libre Graphical Framework）公开
 *                         函数库「Math」分类下 N 次根函数的功能分类与参数域
 *                         （被开方数 + 根次数 两段输入，值 + 有效位 输出），
 *                         只借分类、参数域与命名习惯，算法与实现 100% 自有
 *                         clean-room，不构成衍生作品。
 * 依赖     (Depends)    : 无 DL_ 内部依赖；仅 Standard.library 的 EXP / LN / SQRT
 * 故障码表 (Error codes):
 *   16#0001_011B【信息级】根次数越界（须 1 到 64），返回 0，bValid = FALSE
 *   16#0001_011C【信息级】偶次根负数、入参非有限或结果非有限，返回 0，bValid = FALSE
 * 验收向量 (Acceptance) :
 *   V1 27 的 3 次根 → 3.0（容差 1E-9）
 *   V2 -27 的 3 次根 → -3.0（奇次负数根，符号保留）
 *   V3 -4 的 2 次根 → 0.0，bValid = FALSE，码 011C
 *   V4 16 的 4 次根 → 2.0
 *   V5 根次数 0 → 0.0，码 011B
 *   V6 被开方数 0 → 0.0，bValid = TRUE（不走 LN(0) 路径）
 * 红线自检 (Redline)    : R1 零全局变量表与外部变量引用 ｜ R2 零物理地址直写
 *                         R3 纯 IEC 61131-3 ｜ R4 除零守卫 + 非有限值复检 +
 *                         浮点判零用容差 ｜ R5 全变量中英双语同行注释
 *                         R6 N/A（纯函数无状态机）｜ R7 N/A（无实例调用）
 * 修订历史 (Revision)   :
 *   2026-11-15  v1.0.0  首版入库（Round 10 · Level 1 数学族回补）
 *============================================================================*)

(*==============================================================================
 * 算法推演 (Worked traces)：
 *   推演 1  fValue = 27，nRoot = 3
 *     段 2 根次数 3 在 1 到 64 域内，通过
 *     段 3 入参有限，通过
 *     段 4 绝对值 27 不小于容差，不走零分支
 *     段 5 非负，标记非负，绝对值取 27
 *     段 6 不是一次根、不是二次根、底数不为 1，走对数法：
 *           指数项为 1 除以 3 约 0.3333，自然对数 27 约 3.2958，
 *           二者相乘约 1.0986，取指数得约 3.0
 *     段 7 结果有限，通过
 *     段 8 返回 3.0，有效为真
 *   推演 2  fValue = 负 27，nRoot = 3
 *     段 5 判负成立，根次数为奇数，标记为负，绝对值取 27，余同推演 1
 *     段 6 末段把结果取反，得负 3.0
 *   推演 3  fValue = 负 4，nRoot = 2
 *     段 5 判负成立且根次数为偶数，立即置码 011C 并返回 0，不做任何开方
 *   推演 4  fValue = 0，nRoot = 5
 *     段 4 绝对值小于容差，直接返回 0 且有效为真，绕开对零取对数
 *============================================================================*)

(*==============================================================================
 * 精度与适用域说明 (Accuracy)：
 *   1 二次根走标准库平方根，误差在最低有效位量级；
 *   2 其余次根走「对数加指数」，在双精度下相对误差约 1E-15 量级，
 *     但要求被开方数不为零且根次数不极端大；
 *   3 根次数超过 64 时，底数稍大就会因指数极小而使有效位被吃掉，
 *     故域上限锁在 64，超域一律拒绝而不是硬算；
 *   4 被开方数绝对值超过 1E300 视为溢出，直接拒绝，避免指数运算溢出。
 *============================================================================*)

(*==============================================================================
 * 调用示例 (Instance guide)：
 *   风机相似定律反算转速比（流量与转速成正比，功率与转速三次方成正比）：
 *     fRoot := FC_DL_NthRoot(fValue := fPowerRatio, nRoot := 3);
 *     IF bValid AND (fRoot > 0.0) THEN
 *         fSpeedRatio := fRoot;
 *     END_IF
 *   几何平均（三测点平均直径）：
 *     fGeo := FC_DL_NthRoot(fValue := fA * fB * fC, nRoot := 3);
 *   注意：本件为纯函数，调用后必须判 bValid 再使用返回值；返回 0 既可能是
 *   真实结果（被开方数为零），也可能是域错误，二者只能靠 bValid 与 uErrorId
 *   区分，这是本库对「不返回错误数值冒充结果」红线的具体落地。
 *============================================================================*)

FUNCTION FC_DL_NthRoot : LREAL
VAR_INPUT
    fValue : LREAL := 1.0;   // 被开方数，偶次根要求大于等于 0 [无量纲或工程单位] / Radicand, must be non-negative for even roots
    nRoot  : INT := 2;       // 根次数 n，有效域 1 到 DL_ROOT_MAX（正整数）[次] / Root order, valid 1 to DL_ROOT_MAX
END_VAR
VAR_OUTPUT
    bValid   : BOOL;         // 计算有效（域合法且结果有限）[-] / TRUE when the domain is legal and the result is finite
    uErrorId : UDINT;        // 事件码，0 = 无事件 / Event code, 0 = no event
END_VAR
VAR
    fAbsValue : LREAL;       // 被开方数绝对值，负数路径专用 [无量纲或工程单位] / Absolute value of the radicand
    fResult   : LREAL;       // 计算结果中间量 [无量纲或工程单位] / Result temporaries
    fExpInv   : LREAL;       // 根次数的倒数（如 0.25 对应四次根）[-] / Reciprocal of the root order
    bNegative : BOOL;        // 被开方数是否为负（奇次根取反标志）[-] / TRUE when the radicand is negative
END_VAR
VAR CONSTANT
    DL_ROOT_MIN  : INT   := 1;        // 根次数下限，1 次根等于原值 [次] / Lowest root order, one means identity
    DL_ROOT_MAX  : INT   := 64;       // 根次数上限，超此域对数法精度不可控 [次] / Highest root order
    DL_FLOAT_EPS : LREAL := 1.0E-12;  // 判零与判负容差 [-] / Tolerance for zero and negative tests
    DL_BIG       : LREAL := 1.0E300;  // 非有限值兜底门限 [-] / Magnitude guard for non-finite detection
END_VAR

(*------------------------------------------------------------------------------
 * 段 1｜返回值与标志预置：任何早退路径都要给出确定的 0
 *      Pre-set return value and flags: deterministic zero on every early exit
 *-----------------------------------------------------------------------------*)
FC_DL_NthRoot := 0.0;
bValid        := FALSE;
uErrorId      := 16#0000_0000;
bNegative     := FALSE;

(*------------------------------------------------------------------------------
 * 段 2｜根次数域校验（边界 B1）：必须落在 1 到 64 的闭区间
 *      Root order bounds check (boundary B1)
 *      上限取 64 的工程理由：再大的根次数在单精度输入下有效位已耗尽，
 *      对数法误差会放大到不可接受
 *-----------------------------------------------------------------------------*)
IF (nRoot < DL_ROOT_MIN) OR (nRoot > DL_ROOT_MAX) THEN
    uErrorId := 16#0001_011B;   // 根次数越界，返回 0
    RETURN;
END_IF

(*------------------------------------------------------------------------------
 * 段 3｜入参有限性校验（边界 B2）：NaN 与超大幅值一律拒绝
 *      Input finiteness check (boundary B2): reject NaN and huge magnitudes
 *      NaN 判据用「不等于自身」，是可移植写法，不依赖厂商 ISNAN
 *-----------------------------------------------------------------------------*)
IF (fValue <> fValue) OR (ABS(fValue) > DL_BIG) THEN
    uErrorId := 16#0001_011C;   // 入参非有限
    RETURN;
END_IF

(*------------------------------------------------------------------------------
 * 段 4｜零与近零：直接返回 0，绕开 LN(0) 的负无穷
 *      Zero and near-zero: return 0 directly to bypass LN of zero
 *-----------------------------------------------------------------------------*)
IF ABS(fValue) < DL_FLOAT_EPS THEN
    FC_DL_NthRoot := 0.0;
    bValid        := TRUE;
    RETURN;
END_IF

(*------------------------------------------------------------------------------
 * 段 5｜负数分治（边界 B3）：偶次根无解直接拒绝，奇次根取绝对值后取反
 *      Negative radicand split: even roots are rejected, odd roots keep the sign
 *-----------------------------------------------------------------------------*)
IF fValue < (-1.0 * DL_FLOAT_EPS) THEN
    IF (nRoot MOD 2) = 0 THEN
        uErrorId := 16#0001_011C;   // 偶次根负数，实数域无解，禁止拿绝对值冒充
        RETURN;
    END_IF
    bNegative := TRUE;              // 奇次根：结果保留负号
    fAbsValue := -fValue;
ELSE
    fAbsValue := fValue;
END_IF

(*------------------------------------------------------------------------------
 * 段 6｜主计算：一次根、平方根、底数为一特判，其余走对数法
 *      Main computation: identity, square root and unity shortcuts, then logs
 *      除数 nRoot 已由段 2 保证大于等于 1，不存在除零面
 *-----------------------------------------------------------------------------*)
IF nRoot = DL_ROOT_MIN THEN
    fResult := fAbsValue;                                  // 一次根等于原值
ELSIF (nRoot = 2) AND (NOT bNegative) THEN
    fResult := SQRT(fAbsValue);                            // 平方根走标准库，精度优于对数法
ELSIF ABS(fAbsValue - 1.0) < DL_FLOAT_EPS THEN
    fResult := 1.0;                                        // 底数为 1 时任何次根均为 1
ELSE
    fExpInv := 1.0 / INT_TO_LREAL(nRoot);                  // 根次数倒数，显式类型转换
    fResult := EXP(LN(fAbsValue) / INT_TO_LREAL(nRoot));   // 对数法：e 的 (ln x 除以 n) 次幂
END_IF

IF bNegative THEN
    fResult := -fResult;                                   // 奇次根：符号还原
END_IF

(*------------------------------------------------------------------------------
 * 段 7｜结果有限性复检（边界 B4）：EXP 溢出兜底
 *      Result finiteness recheck (boundary B4): catch exponential overflow
 *-----------------------------------------------------------------------------*)
IF (fResult <> fResult) OR (ABS(fResult) > DL_BIG) THEN
    uErrorId      := 16#0001_011C;   // 结果非有限
    FC_DL_NthRoot := 0.0;
    bValid        := FALSE;
    RETURN;
END_IF

(*------------------------------------------------------------------------------
 * 段 8｜合法收口
 *      Legal close-out
 *-----------------------------------------------------------------------------*)
FC_DL_NthRoot := fResult;
bValid        := TRUE;
END_FUNCTION

(* ---- FC_DL_PercentileLReal.st ---- *)
(*==============================================================================
 * 组件名称 (Component)  : FC_DL_PercentileLReal
 * 所属子库 (Sublibrary) : DL_MathData
 * 当前版本 (Version)    : 1.0.0
 * 分类     (Category)   : 统计函数（Function · Statistics / Pure function）
 * 兼容性   (Platform)   : CODESYS 3.5 / TwinCAT 3 / 汇川 InoProShop / Machine Expert
 *                         仅依赖 Standard.library（LREAL 比较 / 显式类型转换），零厂商方言
 * 功能描述 (Function)   : 对定长样本数组求任意分位值（P0 至 P100），采用业界主流的
 *                         「排序 + 线性插值」口径（R-7 定义，与主流统计库默认一致），
 *                         用于节拍抖动 P95、称重偏差 P99、温度分布 P50 等现场统计判据。
 *                         函数内部完成**拷贝排序**：调用方数组保持原样，与库内就地
 *                         排序件的语义相反，此处刻意如此，见下方不变性声明。
 *
 * 【引脚契约 / Pin contract】
 *   输入 nCount    : INT   — 样本数 [个]，有效域 0 至 64，超上限按 64 截取；
 *   输入 fP        : REAL  — 分位点 [0.0 至 1.0]，0.95 表示 P95，越界钳位；
 *   输入输出 afData: LREAL 数组 [1..64] — 样本数组 [任意工程单位]，
 *                             **只读语义**：函数不写回任何元素，调用方数据帧后不变；
 *   输出 fActualP  : REAL  — 实际生效的分位点（钳位后的值）；
 *   输出 nGuard    : DINT  — 本次排序与拷贝循环的累计次数（防死锁计数，兼作性能诊断）；
 *   输出 bEmpty    : BOOL  — 有效样本为空（或全部非有限 / 排序保护触发），返回 0.0；
 *   输出 uErrorId  : UDINT — 事件码，0 = 无。本件全部码为信息级；
 *   返回  值        : LREAL — 分位值 [与样本同单位]，空集时返回 0.0。
 *
 * 【算法分步 / Algorithm steps（R-7 线性插值口径，写死防漂移）】
 *   ① 样本数闸门：nCount 小于 1 → 空集，返回 0.0、bEmpty 置位、置 0002_000E；
 *      nCount 大于 64 → 只取前 64 个，置 0124（信息级提示，不中断）；
 *   ② 分位点钳位：小于 0 钳到 0，大于 1 钳到 1，非有限（NaN）按 0 处理，置 0124；
 *      fActualP 输出钳位后的实际生效值，供 HMI 显示「实际用的是哪个分位」；
 *   ③ 拷贝筛选取样：把有效样本逐个拷进块内私有数组，**非有限样本直接剔除**
 *      （NaN 参与比较会让整个排序失去传递性，必须前置剔除而不是排序后过滤）；
 *      剔除后为空 → 按空集处理，置 0002_000E；
 *   ④ 插入排序：样本上限 64，插入排序的常数项小于快排且无递归、无栈深风险，
 *      对本规模是最优选择；两层循环均受同一防死锁计数约束；
 *   ⑤ 位置计算：pos = fActualP × (n − 1)，nLo 为 pos 的整数部分（向下取整，
 *      pos 恒非负，截断即向下），fFrac 为小数部分；
 *   ⑥ 插值取值：若 nLo 已到末位则直接取末元素（不外插，P100 恒为最大值）；
 *      否则取第 nLo 与第 nLo+1 个（数组 1 起，故下标分别加 1 与加 2）做线性插值；
 *   ⑦ 结果守卫：插值结果非有限时返回 0.0 并置 0124，绝不把 NaN 交给调用方。
 *
 * 【数组不变性声明 / Array immutability（与就地排序件的语义差异）】
 *   库内排序件（就地快速排序）会改写调用方数组，本件**不会**：全部排序都在块内
 *   私有数组上完成。两种语义同时存在于库内是刻意的——统计取值不应破坏现场数据，
 *   而复用同一份样本做多种统计时更需要原数组保持不变。
 *   代价是每次调用多做一次 64 元素的拷贝，扫描周期量级可忽略。
 *
 * 【为什么本件不调用库内排序件 / Why the sort is inlined】
 *   DL_MathData 层虽然可以依赖本层其他件，但本批六件按要求零互相依赖：
 *   若调用就地快排，则必须先把调用方数组整体备份再回写，既多一次拷贝，
 *   又会在保护触发时留下「部分有序」的中间态，语义反而更差。故内联插入排序。
 *
 * 【边界防错清单 / Boundary guard list】
 *   B1 nCount 小于 1 → 空集返回 0.0、bEmpty 置位、置 0002_000E；
 *   B2 nCount 大于 64 → 截到 64 并置 0124（不越界读取调用方数组）；
 *   B3 fP 越界或非有限 → 钳到 0 或 1，置 0124，继续计算；
 *   B4 样本含 NaN / 无穷 → 剔除该样本；剔除后为空则按空集处理；
 *   B5 排序循环防死锁：拷贝与排序共用 nGuard，超上限即停止、置 bEmpty 并按空集返回，
 *      绝不返回「部分有序」的结果冒充成功；
 *   B6 插值下标双检：nLo 必在 0 至 nN−1 之间，取 nLo+1 与 nLo+2 前先判 nLo+1 是否
 *      越界，越界改取末元素，杜绝数组越界读；
 *   B7 单样本（nCount 为 1）→ pos 恒为 0，直接返回该样本，不外插；
 *   B8 浮点比较全为有序比较（大于 / 小于）；「零个样本」这类判据落在整数域，
 *      浮点判等红线在本件不适用。
 *
 * 【与既有件的职责边界 / Family separation】
 *   FB_DL_SignalStatistics  = 均值 / 方差 / 极值（不含分位）；
 *   FC_DL_QuickSortLReal    = 只排序不取值，且就地改写调用方数组；
 *   本件                    = 排序 + 分位插值，拷贝排序不改调用方数组。
 *   三者互不可替代：要「均值与方差」用统计件，要「有序副本」用排序件，
 *   要「某个分位点上的值」才用本件。
 *
 * 【调用示例 / Call example（仅行注释，不嵌套块注释）】
 *   // 节拍抖动判据：最近 32 个节拍的 P95 超过 12.5 秒即提示瓶颈工位
 *   // fP95 := FC_DL_PercentileLReal(nCount := 32, fP := 0.95,
 *   //          afData := afCycleTime, fActualP => fUsedP, nGuard => nSortCnt,
 *   //          bEmpty => bNoSample, uErrorId => uPctErr);
 *   // IF (NOT bNoSample) AND (fP95 > 12.5) THEN
 *   //     bBottleneckHint := TRUE;
 *   // END_IF
 *
 * 【平台移植注意 / Porting notes】
 *   LREAL 为 64 位浮点，三平台一致；类型转换全部显式写出（REAL 到 LREAL、
 *   LREAL 到 INT），不做隐式提升；插入排序无递归、无栈使用，嵌入式运行时安全；
 *   数组上下界由常量与循环上界双重约束，不依赖动态边界函数。
 *
 * 【工程背景与应用场景 / Background and use cases】
 *   ① 节拍分析：P50 反映典型节拍，P95 反映抖动尾部，两者之差即瓶颈裕度；
 *   ② 称重 / 灌装偏差：P99 用于判定「最差 1 个百分点是否超差」，比均值更贴近验收口径；
 *   ③ 温度分布：多测点 P50 作为炉温代表值，抗单点传感器漂移；
 *   ④ 来料尺寸抽检：P5 与 P95 构成 90 个百分点的居中区间，用于与公差带做对撞判定。
 *
 * 【验收向量 / Acceptance vectors】
 *   V1 中位：样本 1, 2, 3, 4，fP = 0.5 → pos 1.5 → 2 + 0.5 × (3 − 2) = 2.5；
 *   V2 P90：同样本，fP = 0.9 → pos 2.7 → 3 + 0.7 × (4 − 3) = 3.7；
 *   V3 单样本：样本 7.5，fP = 0.9 → 7.5（pos 为 0，不外插）；
 *   V4 越界钳位：fP = 1.5、样本 1, 2, 3, 4 → fActualP 1.0、返回 4.0、置 0124；
 *   V5 空集：nCount 为 0 → 返回 0.0、bEmpty 置位、置 0002_000E；
 *   V6 输入不变：样本 4, 1, 3, 2，fP = 0.5 → 返回 2.5，且调用方数组帧后仍为原序。
 *
 * 【事件码表 / Event code table（全部信息级，不置报警位）】
 *   16#0001_0124  分位点或样本数越界已钳位 / 非有限样本已剔除 / 结果非有限已回退；
 *   16#0002_000E  有效样本为空（含全部非有限与排序保护触发），返回 0.0。
 *
 * 修订历史 (Revision)   :
 *   2026-11-15  v1.0.0  首版落盘（Round 11 · 泳道 A · LGF Math 组）
 *============================================================================*)
FUNCTION FC_DL_PercentileLReal : LREAL
VAR_INPUT
    nCount : INT;                          // 样本数 [个]，有效域 0 至 64 / Sample count [pcs], valid range 0 to 64
    fP     : REAL;                         // 分位点 [0.0 至 1.0]，0.95 即 P95 / Percentile [0.0 to 1.0], 0.95 means P95
END_VAR
VAR_IN_OUT
    afData : ARRAY[1..64] OF LREAL;        // 样本数组 [工程单位]，只读语义，块内拷贝 / Sample array [EU], read-only, copied internally
END_VAR
VAR_OUTPUT
    fActualP : REAL;                       // 实际生效的分位点，越界已钳位 / Effective percentile after clamping
    nGuard   : DINT;                       // 循环累计次数，防死锁兼性能诊断 / Loop counter for guard and diagnostics
    bEmpty   : BOOL;                       // 有效样本为空，返回 0.0 / Empty valid sample set, returns 0.0
    uErrorId : UDINT;                      // 事件码，0 = 无 / Event code, 0 = none
END_VAR
VAR
    afSorted : ARRAY[1..64] OF LREAL;      // 块内私有排序数组，不触碰调用方 / Private sorted array, the caller array is untouched
    nUsable  : INT;                        // 本拍可读样本上界 [个] / Readable sample upper bound of this scan [pcs]
    nN       : INT;                        // 剔除非有限后的有效样本数 [个] / Effective sample count after filtering [pcs]
    nI       : INT;                        // 外层索引 / Outer index
    nJ       : INT;                        // 内层回退索引 / Inner shift index
    fKey     : LREAL;                      // 当前插入键值 [工程单位] / Current insertion key [EU]
    bShift   : BOOL;                       // 内层回退继续标志 / Inner shift continues flag
    bSortOk  : BOOL;                       // 排序完整完成标志 / Sort completed flag
    fPos     : LREAL;                      // 分位在样本序列上的位置 [-] / Percentile position in the sample sequence [-]
    nLo      : INT;                        // 位置整数部分（截断） / Integer part of the position, truncated
    fFrac    : LREAL;                      // 位置小数部分 [-] / Fractional part of the position [-]
    fLo      : LREAL;                      // 插值下样本值 [工程单位] / Lower interpolation sample [EU]
    fHi      : LREAL;                      // 插值上样本值 [工程单位] / Upper interpolation sample [EU]
    fResult  : LREAL;                      // 插值结果工作副本 [工程单位] / Working copy of the interpolation result [EU]
END_VAR
VAR CONSTANT
    DL_SAMPLE_MAX : INT   := 64;           // 样本上限 [个]，与数组维度一致 / Sample upper bound [pcs], matches the array
    DL_GUARD_MAX  : DINT  := 100000;       // 循环防死锁上限 [次] / Loop guard limit [count]
    DL_FLOAT_EPS  : REAL  := 1.0E-6;       // 浮点容差 [-] / Float epsilon [-]
    DL_LL_EPS     : LREAL := 1.0E-9;       // 长浮点容差 [-] / Long-real epsilon [-]
    DL_P_MIN      : REAL  := 0.0;          // 分位点下界 / Percentile lower bound
    DL_P_MAX      : REAL  := 1.0;          // 分位点上界 / Percentile upper bound
    DL_LL_ZERO    : LREAL := 0.0;          // 长浮点零值 / Long-real zero
    DL_LL_ONE     : LREAL := 1.0;          // 长浮点一值，位置计算的减数 / Long-real one, used in the position formula
    DL_INF_LIM    : LREAL := 1.0E300;      // 非有限值判据阈值 / Non-finite threshold
    DL_ERR_CLAMP  : UDINT := 16#0001_0124; // 钳位与剔除的信息级码 / Info code for clamping and filtering
    DL_ERR_EMPTY  : UDINT := 16#0002_000E; // 有效样本为空的信息级码 / Info code for an empty valid sample set
END_VAR

(*------------------------------------------------------------------------------
 * 段 1｜返回值与输出预置（函数必须先给出安全返回值）
 *      Preset the return value and the outputs
 *   返回值预置 0.0、bEmpty 预置假：只有明确判定为空集时才置真，避免误报。
 *-----------------------------------------------------------------------------*)
FC_DL_PercentileLReal := DL_LL_ZERO;       // 返回值预置 0（Return preset to zero）
fActualP  := DL_P_MIN;                     // 生效分位点预置下界（Effective percentile preset）
nGuard    := 0;                            // 循环计数清零（Loop guard cleared）
bEmpty    := FALSE;                        // 空集标志预置假（Empty flag preset false）
uErrorId  := 16#0000_0000;                 // 事件码预清零（Event code preset to zero）
bSortOk   := TRUE;                         // 排序完成标志预置真（Sort flag preset true）
nN        := 0;                            // 有效样本数预置 0（Effective count preset）
nUsable   := 0;                            // 可读样本数预置 0（Readable count preset）
fResult   := DL_LL_ZERO;                   // 结果副本预置 0（Result working copy preset）

(*------------------------------------------------------------------------------
 * 段 2｜样本数闸门与可读上界（边界 B1 / B2）
 *      Sample count gate and the readable upper bound
 *   上界同时受「调用方声明数」与「数组容量」双重约束：取小者，
 *   任何情况下都不会读出数组之外。
 *-----------------------------------------------------------------------------*)
IF nCount < 1 THEN                         // 无样本（No samples declared）
    bEmpty   := TRUE;                      // 置空集标志（Raise the empty flag）
    uErrorId := DL_ERR_EMPTY;              // 置空集信息码（Raise the empty info code）
    RETURN;                                // 早退，返回值保持 0.0（Early exit, return stays zero）
END_IF

nUsable := nCount;                         // 可读上界先取声明数（Readable bound takes the declared count）
IF nUsable > DL_SAMPLE_MAX THEN            // 超数组容量（Above the array capacity）
    nUsable  := DL_SAMPLE_MAX;             // 截到容量，杜绝越界读（Truncate to the capacity）
    uErrorId := DL_ERR_CLAMP;              // 置截断信息码（Raise the truncation info code）
END_IF

(*------------------------------------------------------------------------------
 * 段 3｜分位点钳位（边界 B3）
 *      Percentile clamping
 *   次序写死：先判上越界、再判下越界、最后判非有限（NaN 与两个有序比较都为假）。
 *   非有限按 0 处理而不是按 1 处理：0 分位取最小值，属保守回退。
 *-----------------------------------------------------------------------------*)
fActualP := fP;                            // 生效分位点先接管输入（Take the input percentile）
IF fP > DL_P_MAX THEN                      // 上越界（Above the upper bound）
    fActualP := DL_P_MAX;                  // 钳到 1（Clamp to one）
    uErrorId := DL_ERR_CLAMP;              // 置钳位信息码（Raise the clamp info code）
ELSIF fP < DL_P_MIN THEN                   // 下越界（Below the lower bound）
    fActualP := DL_P_MIN;                  // 钳到 0（Clamp to zero）
    uErrorId := DL_ERR_CLAMP;              // 置钳位信息码（Raise the clamp info code）
ELSIF NOT ((fP <= DL_P_MAX) AND (fP >= DL_P_MIN)) THEN   // 非有限值，NaN 落入此支（Not finite, NaN path）
    fActualP := DL_P_MIN;                  // 保守按 0 分位（Fall back to the zero percentile）
    uErrorId := DL_ERR_CLAMP;              // 置钳位信息码（Raise the clamp info code）
END_IF

(*------------------------------------------------------------------------------
 * 段 4｜拷贝取样并剔除非有限样本（边界 B4）
 *      Copy the samples and filter out the non-finite ones
 *   NaN 参与比较会让排序失去传递性，必须在排序**之前**剔除，而不是排完再过滤。
 *-----------------------------------------------------------------------------*)
FOR nI := 1 TO nUsable DO                  // 只遍历可读区间（Iterate the readable range only）
    nGuard := nGuard + 1;                  // 拷贝循环同样计入防死锁（Counted by the guard）
    IF (afData[nI] <= DL_INF_LIM) AND (afData[nI] >= -DL_INF_LIM) THEN   // 有限样本（Finite sample）
        nN := nN + 1;                      // 有效样本数加 1（Effective count increments）
        afSorted[nN] := afData[nI];        // 拷进私有数组，调用方数组只读（Copy into the private array）
    ELSE                                   // 非有限样本（Non-finite sample）
        uErrorId := DL_ERR_CLAMP;          // 置剔除信息码（Raise the filtering info code）
    END_IF
END_FOR

IF nN < 1 THEN                             // 剔除后无有效样本（No effective sample left）
    bEmpty   := TRUE;                      // 置空集标志（Raise the empty flag）
    uErrorId := DL_ERR_EMPTY;              // 空集码覆盖钳位码，语义优先（The empty code wins）
    RETURN;                                // 早退，返回值保持 0.0（Early exit, return stays zero）
END_IF

(*------------------------------------------------------------------------------
 * 段 5｜插入排序（边界 B5：两层循环共用防死锁计数）
 *      Insertion sort with a shared guard counter
 *   样本不超过 64，插入排序常数项小、无递归、无栈深风险，对本规模最优；
 *   超出防护上限即判定排序未完成，绝不把「部分有序」冒充成功。
 *-----------------------------------------------------------------------------*)
FOR nI := 2 TO nN DO                       // 从第二个元素起逐个插入（Insert from the second element）
    IF nGuard > DL_GUARD_MAX THEN          // 早期熔断，避免无谓空转（Early trip to avoid spinning）
        bSortOk := FALSE;                  // 标记未完成（Mark as incomplete）
        EXIT;                              // 跳出外层循环（Leave the outer loop）
    END_IF

    fKey   := afSorted[nI];                // 当前待插入键值（Current insertion key）
    nJ     := nI - 1;                      // 从已排序区末位开始回退（Start from the sorted tail）
    bShift := TRUE;                        // 回退标志置真（Shift flag set）

    WHILE bShift AND (nJ >= 1) DO          // 回退直到找到插入位（Shift until the slot is found）
        nGuard := nGuard + 1;              // 内层循环计入防死锁（Counted by the guard）
        IF nGuard > DL_GUARD_MAX THEN      // 触顶熔断（Guard exhausted）
            bShift  := FALSE;              // 停止回退（Stop shifting）
            bSortOk := FALSE;              // 标记未完成（Mark as incomplete）
        ELSIF afSorted[nJ] > fKey THEN     // 前一个更大，后移一格（Shift one slot right）
            afSorted[nJ + 1] := afSorted[nJ];
            nJ := nJ - 1;                  // 索引回退（Index steps back）
        ELSE                               // 找到插入位（Insertion slot found）
            bShift := FALSE;               // 停止回退（Stop shifting）
        END_IF
    END_WHILE

    afSorted[nJ + 1] := fKey;              // 键值落位，nJ 恒非负故下标合法（Place the key, index stays valid）
END_FOR

IF NOT bSortOk THEN                        // 排序未完成，结果不可信（Sort incomplete, result untrusted）
    bEmpty   := TRUE;                      // 按空集处理，绝不返回半成品（Treat as empty, never return a partial result）
    uErrorId := DL_ERR_EMPTY;              // 置空集信息码（Raise the empty info code）
    RETURN;                                // 早退，返回值保持 0.0（Early exit, return stays zero）
END_IF

(*------------------------------------------------------------------------------
 * 段 6｜位置计算（R-7 口径：pos = P × (n − 1)）
 *      Position computation
 *   pos 恒非负，故 LREAL 到 INT 的截断转换等价于向下取整，无需额外取整函数。
 *-----------------------------------------------------------------------------*)
fPos  := REAL_TO_LREAL(fActualP) * (INT_TO_LREAL(nN) - DL_LL_ONE);   // 位置 = P 乘（n 减 1）（Position formula）
nLo   := LREAL_TO_INT(fPos);               // 整数部分，pos 非负故截断即向下（Truncation equals floor here）
fFrac := fPos - INT_TO_LREAL(nLo);         // 小数部分（Fractional part）

IF nLo < 0 THEN                            // 理论上不可达的兜底（Unreachable fallback）
    nLo := 0;                              // 索引归零（Index reset）
    fFrac := DL_LL_ZERO;                   // 小数部分归零（Fraction reset）
END_IF
IF nLo > (nN - 1) THEN                     // 上限兜底（Upper fallback）
    nLo := nN - 1;                         // 钳到末位（Clamp to the last slot）
    fFrac := DL_LL_ZERO;                   // 小数部分归零（Fraction reset）
END_IF

(*------------------------------------------------------------------------------
 * 段 7｜线性插值取值（边界 B6 / B7：下标双检，末位不外插）
 *      Linear interpolation with double index checks
 *   数组 1 起：第 k 个样本（0 起计）位于下标 k+1，故下样本取 nLo+1、上样本取 nLo+2。
 *-----------------------------------------------------------------------------*)
IF (nLo + 1) >= nN THEN                    // 已到末位，直接取最大样本（Last slot, take the maximum）
    fResult := afSorted[nN];               // 不外插，P100 恒为最大值（No extrapolation）
ELSE                                       // 需要插值（Interpolation required）
    fLo := afSorted[nLo + 1];              // 下样本（Lower sample）
    fHi := afSorted[nLo + 2];              // 上样本，下标已由上一支保证不越界（Upper sample, bounds proven）
    fResult := fLo + fFrac * (fHi - fLo);  // 线性插值（Linear interpolation）
END_IF

(*------------------------------------------------------------------------------
 * 段 8｜结果守卫（边界 B8）
 *      Post guard on the interpolation result
 *   非有限结果一律回退 0.0：统计值的下游多为比较与报警，NaN 会在那里静默失效。
 *-----------------------------------------------------------------------------*)
IF NOT ((fResult <= DL_INF_LIM) AND (fResult >= -DL_INF_LIM)) THEN   // 结果非有限（Non-finite result）
    fResult   := DL_LL_ZERO;               // 回退 0（Fall back to zero）
    uErrorId  := DL_ERR_CLAMP;             // 置回退信息码（Raise the fallback info code）
END_IF

FC_DL_PercentileLReal := fResult;          // 结果落位（Place the result）
END_FUNCTION

(* ---- FC_DL_RandomNext.st ---- *)
(*==============================================================================
 * 组件名称 (Component)  : FC_DL_RandomNext
 * 所属子库 (Sublibrary) : DL_MathData
 * 当前版本 (Version)    : 1.0.0
 * 分类     (Category)   : 随机序列函数（Function · Math / Test stimulus）
 * 兼容性   (Platform)   : CODESYS 3.5 / TwinCAT 3 / 汇川 InoProShop / Machine Expert
 *                         仅依赖 Standard.library（UDINT 乘加 / 显式类型转换），零厂商方言
 * 功能描述 (Function)   : 线性同余（乘加型）伪随机序列的**单步递推**。给定当前
 *                         种子返回 [0, 1) 区间的均匀分布随机数与**新种子**，函数
 *                         内部不保存任何状态：调用方只需把 uNextSeed 回灌下一拍，
 *                         即可得到「可复现、可回溯、可插入断点」的确定序列。
 *                         用于通讯压力测试、仿真激励、算法自检与随机抽样验证。
 *
 * 【引脚契约 / Pin contract】
 *   输入 uSeed      : UDINT — 当前种子 [cnt]，首次调用由调用方给定任意值；
 *   输入 bReseed    : BOOL  — TRUE 时强制改用内置默认种子（可复现基线）；
 *   输出 uNextSeed  : UDINT — 下一拍应回灌的种子 [cnt]；
 *   输出 bZeroSeed  : BOOL  — 本次输入种子为 0，已置提示位（见下方勘误声明）；
 *   输出 bSat      : BOOL  — 结果被钳到 1.0 减容差，保证半开区间；
 *   输出 uErrorId  : UDINT — 事件码，0 = 无。本件全部码为信息级；
 *   返回  值        : REAL  — [0, 1) 均匀分布随机数。
 *
 * 【递推式与参数 / Recurrence and parameters】
 *   uNextSeed = uSeed × 1664525 + 1013904223（以 2 的 32 次方为模，无符号自然回绕）
 *   参数取自《Numerical Recipes》公开推荐的乘加型同余参数：
 *   周期为 2 的 32 次方（全周期），高 16 位统计质量良好，足够测试激励使用。
 *   本件**不显式取模**：无符号 32 位乘加的溢出回绕在三平台语义一致，
 *   显式取模反而会引入「有符号 / 无符号取模行为差异」这一类历史坑。
 *
 * 【可复现性承诺 / Reproducibility contract】
 *   同一 (uSeed, bReseed) 输入组合，在任何扫描周期、任何平台、任何时刻调用，
 *   返回值与 uNextSeed 完全一致；不存在「上电时间参与」或「内部状态漂移」。
 *   由此得到两条可用的自检关系：
 *     R1 反向复算：FLOOR(返回值 / 2.3283064E-10) 等于 uNextSeed（容差内）；
 *     R2 序列复现：把 uNextSeed 回灌，第二次调用的结果与首次运行同序号一致。
 *
 * 【归一与半开区间 / Normalisation and the half-open interval】
 *   返回值 = uNextSeed × 2.3283064E-10（即乘以 2 的 32 次方的倒数）。
 *   由于 REAL 只有 24 位尾数，极大种子在归一乘之后可能被舍入到 1.0，
 *   故在后置守卫里把「大于等于 1.0」的结果钳到 1.0 减容差并置 bSat，
 *   以此**硬保证**返回值落在 [0, 1) 半开区间——这是调用方做数组下标
 *   （乘以容量后取整）时不会越界的唯一前提。
 *
 * 【对规格原文的一处勘误 / Erratum on the specification】
 *   规格原文称「0 在乘法型同余中是吸收态，需替换为默认种子」。经复核：本件采用
 *   **增量非零**的乘加型（增量 1013904223 为奇数），零种子经一次递推即得增量本身，
 *   随后立即脱离零，并不是吸收态；若强行替换为默认种子，则与同一规格给出的
 *   验收向量「零种子 → 新种子 = 1013904223」直接矛盾。故本实现取：
 *   零种子**按原值参与递推**，同时置 bZeroSeed 供现场识别「种子未初始化」，
 *   序列既满足向量，也不产生退化。此为刻意决策，不是遗漏。
 *
 * 【边界防错清单 / Boundary guard list】
 *   B1 乘子被工具链改写为 0（理论上不可达）→ 回退到增量常数（奇数非零），
 *      置 0123，保证任何情况下序列不退化；
 *   B2 种子为 0 → 按原值递推并置 bZeroSeed（见勘误声明），不产生常数列；
 *   B3 重播种（bReseed TRUE）→ 强制从默认种子起步，优先级高于零种子提示；
 *   B4 归一结果舍入到 1.0 → 钳到 1.0 减容差并置 bSat，保证半开区间；
 *   B5 归一结果为负（理论上不可达）→ 钳到 0.0，保证下界；
 *   B6 全件无除法（用乘法倒数代替）、无数组、无循环，不存在除零、越界、死循环；
 *   B7 浮点比较只做区间与下界判断（有序比较），唯一「等于 0」的判据落在
 *      UDINT 域（整数判等合法），浮点判等红线在本件不适用。
 *
 * 【与既有件的职责边界 / Family separation】
 *   FB_DL_SineGenerator / FB_DL_SawtoothGenerator / FB_DL_PulseGenerator
 *   = 确定性**波形**发生器（周期、相位、幅值可调，输出形状固定）；
 *   本件 = **伪随机**序列且**无状态**（不占实例内存、可重入、可回溯）。
 *   波形件给「可预期的激励」，本件给「不可预期但可复现的激励」，用途正交。
 *
 * 【调用示例 / Call example（仅行注释，不嵌套块注释）】
 *   // 通讯压力测试：每拍生成一个随机报文号，种子由静态变量持有
 *   // fRand := FC_DL_RandomNext(uSeed := uMySeed, bReseed := bTestRestart,
 *   //          uNextSeed => uMySeed, bZeroSeed => bSeedBad,
 *   //          bSat => bRandSat, uErrorId => uRandErr);
 *   // uMsgNo := REAL_TO_UDINT(fRand * 1000.0);   // 0 ~ 999 的报文号
 *
 * 【平台移植注意 / Porting notes】
 *   UDINT 乘加溢出回绕在三平台一致；UDINT 到 REAL 的转换按「显式转换」写出，
 *   不做隐式提升；本件不依赖任何随机数系统函数（平台各有方言，且不可复现）。
 *
 * 【工程背景与应用场景 / Background and use cases】
 *   ① 通讯压力测试：随机长度、随机间隔的报文灌注，压出缓冲区边界缺陷；
 *   ② 仿真激励：给滤波器与统计件灌随机序列，验证极值与分位计算；
 *   ③ 算法自检：同一种子重跑同一序列，比对两次运行结果是否逐位一致；
 *   ④ 抽样巡检：从合格批次里随机抽检，种子留档后可完全复现抽检名单。
 *
 * 【局限与误用提示 / Limitations and misuse】
 *   ① 本件是**测试激励级**序列：低位相关性明显，禁止用于安全相关抽样（如安全
 *      功能抽检名单）、禁止用于加密与鉴权、禁止用于需要统计独立性的 A/B 分流；
 *   ② 序列周期为 2 的 32 次方，长时间高频调用后会出现重复，压力测试可接受，
 *      长周期仿真应由调用方按批次换种子；
 *   ③ 本件不保存状态：调用方若忘记回灌 uNextSeed，每拍都会得到同一个数，
 *      这一类「序列卡死」不是本件故障，排查时先看种子是否回灌；
 *   ④ 需并行多路序列时，各路给不同初值种子即可，本件无共享状态、无互斥需求。
 *
 * 【验收向量 / Acceptance vectors】
 *   V1 零种子：uSeed = 0 → uNextSeed = 1013904223、返回值约 0.2360680、bZeroSeed；
 *   V2 满量程种子：uSeed = 16#FFFF_FFFF → uNextSeed = 1012239698、返回值约 0.2356716；
 *   V3 确定性：同一种子连调两次（第二次回灌 uNextSeed），序列与前次运行一致；
 *   V4 半开区间：任取 1000 个种子，返回值全部满足 0.0 至 1.0 的左闭右开；
 *   V5 重播种：bReseed TRUE 时无论 uSeed 为何，uNextSeed 恒为默认种子的首步结果。
 *   V6 参数退化：把乘子视为 0 的损坏场景 → 回退后序列仍逐拍变化、uErrorId 0123。
 *
 * 【事件码表 / Event code table（全部信息级，不置报警位）】
 *   16#0001_0123  递推参数被改写为退化值，已回退到保底常数（保护性提示）。
 *
 * 修订历史 (Revision)   :
 *   2026-11-15  v1.0.0  首版落盘（Round 11 · 泳道 A · LGF Math 组）
 *============================================================================*)
FUNCTION FC_DL_RandomNext : REAL
VAR_INPUT
    uSeed    : UDINT;                      // 当前种子 [cnt]，首次调用任意值 / Current seed [cnt], any value on the first call
    bReseed  : BOOL;                       // TRUE 时强制从默认种子起步 / TRUE forces the default seed
END_VAR
VAR_OUTPUT
    uNextSeed : UDINT;                     // 下一拍应回灌的种子 [cnt] / Seed to feed back on the next call [cnt]
    bZeroSeed : BOOL;                      // 输入种子为 0 的提示位 / Notice flag for a zero input seed
    bSat      : BOOL;                      // 结果已钳到上界容差内 / Result clamped inside the upper bound
    uErrorId  : UDINT;                     // 事件码，0 = 无 / Event code, 0 = none
END_VAR
VAR
    _uWork   : UDINT;                      // 本次实际参与递推的种子 [cnt] / Seed actually used by the recurrence [cnt]
    _uMul    : UDINT;                      // 工作乘子，含退化回退 / Working multiplier with the fallback
    _uInc    : UDINT;                      // 工作增量，含退化回退 / Working increment with the fallback
    _fOut    : REAL;                       // 归一后的随机数 [-] / Normalised random number [-]
END_VAR
VAR CONSTANT
    DL_LCG_MUL      : UDINT := 1664525;        // 乘子，Numerical Recipes 公开参数 / Multiplier from the Numerical Recipes parameters
    DL_LCG_INC      : UDINT := 1013904223;     // 增量，奇数保证全周期 / Increment, odd ensures a full period
    DL_SEED_DEFAULT : UDINT := 16#0000_0001;   // 默认种子，重播种基线与零种子回退 / Default seed for reseeding and fallback
    DL_RAND_SCALE   : REAL  := 2.3283064E-10;  // 2 的 32 次方倒数，归一因子 / Reciprocal of two to the thirty-second power
    DL_FLOAT_EPS    : REAL  := 1.0E-6;         // 上界保护容差 / Upper-bound guard epsilon
    DL_ONE          : REAL  := 1.0;            // 半开区间上界 / Upper bound of the half-open interval
    DL_RAND_ZERO    : REAL  := 0.0;            // 半开区间下界 / Lower bound of the half-open interval
    DL_ERR_PARAM    : UDINT := 16#0001_0123;   // 递推参数退化回退的信息级码 / Info code for the degenerate parameter fallback
END_VAR

(*------------------------------------------------------------------------------
 * 段 1｜返回值与输出预置（函数必须先给出安全返回值）
 *      Preset the return value and the outputs
 *   返回值预置 0.0：早退路径一律给下界值，绝不给未初始化的中间量。
 *-----------------------------------------------------------------------------*)
FC_DL_RandomNext := DL_RAND_ZERO;          // 返回值预置 0（Return preset to zero）
uNextSeed := 0;                            // 新种子预置 0，段 4 覆盖（Next seed preset, overwritten in stage 4）
bZeroSeed := FALSE;                        // 零种子提示位预置（Zero-seed notice preset）
bSat      := FALSE;                        // 上限钳位标志预置（Upper clamp flag preset）
uErrorId  := 16#0000_0000;                 // 事件码预清零（Event code preset to zero）

(*------------------------------------------------------------------------------
 * 段 2｜递推参数的完整性校验（边界 B1）
 *      Integrity check of the recurrence parameters
 *   乘子为 0 会让序列退化成常数列（每拍都等于增量），这是唯一致命的参数损坏；
 *   出现时回退到增量常数（奇数且非零），并置信息码留痕，绝不静默继续。
 *-----------------------------------------------------------------------------*)
_uMul := DL_LCG_MUL;                       // 乘子工作副本接管常数（Multiplier working copy）
_uInc := DL_LCG_INC;                       // 增量工作副本接管常数（Increment working copy）

IF _uMul = 0 THEN                          // 乘子被改写为 0，序列将退化（Degenerate multiplier）
    _uMul    := DL_LCG_INC;                // 回退到增量常数，保底非零（Fall back to the non-zero increment）
    uErrorId := DL_ERR_PARAM;              // 置参数回退信息码（Raise the parameter fallback info code）
END_IF
IF _uInc = 0 THEN                          // 增量为 0 时退化为纯乘法型（Zero increment degenerates to a pure multiplier）
    _uInc    := DL_LCG_MUL;                // 回退到乘子常数，保底非零（Fall back to the non-zero multiplier）
    uErrorId := DL_ERR_PARAM;              // 置参数回退信息码（Raise the parameter fallback info code）
END_IF

(*------------------------------------------------------------------------------
 * 段 3｜种子选择（边界 B2 / B3：重播种优先，零种子只提示不替换）
 *      Seed selection, reseed wins, a zero seed is only flagged
 *   口径见头注释的勘误声明：零种子按原值参与递推，仅置提示位。
 *-----------------------------------------------------------------------------*)
IF bReseed THEN                            // 重播种请求（Reseed requested）
    _uWork    := DL_SEED_DEFAULT;          // 强制从默认种子起步（Start from the default seed）
    bZeroSeed := FALSE;                    // 重播种时不再提示零种子（No zero-seed notice on a reseed）
ELSE                                       // 常规递推（Regular recurrence）
    _uWork := uSeed;                       // 种子原值接管（Take the input seed as-is）
    IF uSeed = 0 THEN                      // 种子为 0，提示未初始化（Zero seed noticed）
        bZeroSeed := TRUE;                 // 置提示位（Raise the notice flag）
    END_IF
END_IF

(*------------------------------------------------------------------------------
 * 段 4｜单步递推（模 2 的 32 次方，无符号自然回绕，不显式取模）
 *      Single-step recurrence with natural 32-bit wraparound
 *   先乘后加，全程 UDINT 域：回绕由类型宽度自然完成，跨平台一致。
 *-----------------------------------------------------------------------------*)
uNextSeed := _uWork * _uMul + _uInc;       // 递推一步，新种子（One recurrence step, the next seed）

(*------------------------------------------------------------------------------
 * 段 5｜归一化（半开区间由后置守卫硬保证）
 *      Normalisation, the half-open interval is enforced by the guards below
 *   用乘法倒数代替除法：既避开除零，也避开「除以 2 的 32 次方」的精度损失。
 *-----------------------------------------------------------------------------*)
_fOut := UDINT_TO_REAL(uNextSeed) * DL_RAND_SCALE;   // 显式转换后乘以归一因子（Explicit cast then scale）
FC_DL_RandomNext := _fOut;                 // 结果先行落位（Result placed first）

(*------------------------------------------------------------------------------
 * 段 6｜后置守卫（边界 B4 / B5）
 *      Post guards on the returned value
 *   REAL 尾数 24 位，极大种子归一后可能被舍入到 1.0：钳到 1.0 减容差并置 bSat，
 *   这是调用方「乘以容量后取整」不越界的唯一前提。
 *-----------------------------------------------------------------------------*)
IF FC_DL_RandomNext >= DL_ONE THEN         // 舍入触及上界（Rounded up to the bound）
    FC_DL_RandomNext := DL_ONE - DL_FLOAT_EPS;  // 钳到上界内侧（Clamp inside the bound）
    bSat := TRUE;                          // 置钳位标志（Raise the clamp flag）
END_IF

IF FC_DL_RandomNext < DL_RAND_ZERO THEN    // 结果低于下界，理论上不可达（Below the bound, unreachable）
    FC_DL_RandomNext := DL_RAND_ZERO;      // 钳到下界（Clamp to the lower bound）
END_IF
END_FUNCTION
